REGION Network 6: Span Adjustment
   // Zero adjustment has to be performed prior to this linearity adjustment procedure.
   // 
   // 1. Specify how many linearity adjustment points to be performed by loading interger 0, 1, 2 or 3 into LinearityRange (0 for 2 points, 1 for 3 points, 2 for 4 points and 3 for 5 points). Please be noted that the earlier performed zero adjustment point is considered as the first adjustment point (Point #1).
   // 
   // 2. Configure all the adjustment weight values into xLow, Low, Middle and High (for e.g. 5-point adjustment requires all 4 weights: High, Middle, Low and xLow; 3-point requires High and Middle; 2-point only requies High as the 1st point is the zero reference)
   // 
   // 3. Make sure the Linearity Range parameter and all the adjustment weight values are configured correctly before starting the adjustment process. Invalid or incomplete parameters will cause the Function Block to turn on the Error output bit.
   // 
   // 4. Trigger ON  Input Start bit to start the span adjustment. This Start bit will be turned off by the Function Block upon completion/ cancellation or error condition. 
   // 
   // 5. Once started, CurrentPoint shows the current linearity point to be adjusted; CurrentWeight shows current adjustment weight to be loaded onto the scale. The LoadWeight output bit will be set ON to request for new adjustment weight. 
   // 
   // 6. After loading the new adjustment weight, acknowledge this by triggering the ConfirmWeight parameter (boolean) ON. The Function Block will then proceed to the next adjustment point and turn off this ConfirmWeight bit.
   // 
   // 7. Output bit - Process signifies that the adjustment of current point is in process.
   // 
   // 8. Input Parameter Bit Cancel is used to cancel/ abort the adjustment process
   RUNG wire#powerrail
      "SAI_IND_SpanAdjust_DB"(ID := "IND360~Head", Hi_Weight := "SAI_IND_SpanAdjust_DB".Hi_Weight, Mid_Weight := "SAI_IND_SpanAdjust_DB".Mid_Weight, Low_Weight := "SAI_IND_SpanAdjust_DB".Low_Weight, xLow_Weight := "SAI_IND_SpanAdjust_DB".xLow_Weight, LinearityRange := "SAI_IND_SpanAdjust_DB".LinearityRange, Start := "SAI_IND_SpanAdjust_DB".Start, ConfirmWeight := "SAI_IND_SpanAdjust_DB".ConfirmWeight, Cancel := "SAI_IND_SpanAdjust_DB".Cancel, CurrentPoint => "SAI_IND_SpanAdjust_DB".CurrentPoint, CurrentWeight => "SAI_IND_SpanAdjust_DB".CurrentWeight, LoadWeight => "SAI_IND_SpanAdjust_DB".LoadWeight, Process => "SAI_IND_SpanAdjust_DB".Process, Done => "SAI_IND_SpanAdjust_DB".Done, Error => "SAI_IND_SpanAdjust_DB".Error, Cancelled => "SAI_IND_SpanAdjust_DB".Cancelled)
   END_RUNG
   // the same network as SCL:
   "SAI_IND_SpanAdjust_DB"(ID := "IND360~Head",   // "SAI_IND_SpanAdjust"
                           Hi_Weight := "SAI_IND_SpanAdjust_DB".Hi_Weight,
                           Mid_Weight := "SAI_IND_SpanAdjust_DB".Mid_Weight,
                           Low_Weight := "SAI_IND_SpanAdjust_DB".Low_Weight,
                           xLow_Weight := "SAI_IND_SpanAdjust_DB".xLow_Weight,
                           LinearityRange := "SAI_IND_SpanAdjust_DB".LinearityRange,
                           Start := "SAI_IND_SpanAdjust_DB".Start,
                           ConfirmWeight := "SAI_IND_SpanAdjust_DB".ConfirmWeight,
                           Cancel := "SAI_IND_SpanAdjust_DB".Cancel,
                           CurrentPoint => "SAI_IND_SpanAdjust_DB".CurrentPoint,
                           CurrentWeight => "SAI_IND_SpanAdjust_DB".CurrentWeight,
                           LoadWeight => "SAI_IND_SpanAdjust_DB".LoadWeight,
                           Process => "SAI_IND_SpanAdjust_DB".Process,
                           Done => "SAI_IND_SpanAdjust_DB".Done,
                           Error => "SAI_IND_SpanAdjust_DB".Error,
                           Cancelled => "SAI_IND_SpanAdjust_DB".Cancelled);
END_REGION

REGION Network 7: CalFree Adjustment
   // CalFree is a method of analog scale adjustment without using test weights. It takes the factory calibrated load cell Rated Output (mV/ Vexc.) and user defined scale capacity to build a linear loading curve.
   // This method is usually applied to huge capacity scales in which calibration with test weights or other material is not feasible at all. 
   // 
   // For Powercell scale, please use the CalFree+ Function Block instead.
   // 
   // 1. Write in.. 
   // (a) CalFree Scale Capacity (Index 0x401A), 
   // (b) CalFree Scale unit (Index 0x401C, Decimal 0 - gram; Decimal 1 - KG; Decimal 2 - Pounds) and 
   // (c) Load Cells' averaged Rated Output (Index 0x401D, in mV/V)
   // **Make sure the transmitter's scale capacity has already been configured to the same value as CalFree Capacity prior to this CalFree adjustment.
   // 
   // 2. Trigger Input bit Start for CalFree adjustment (Index 0x401A)
   // 
   // 3. Output bit Done will be turned ON after successful completion of the process
   // Error output bit will be turned ON if there is an error during the adjustment process
   RUNG wire#powerrail
      "SAI_IND_CalFree_DB"(ID := "IND360~Head", RatedCapacity := "SAI_IND_CalFree_DB".RatedCapacity, Unit := "SAI_IND_CalFree_DB".Unit, RatedOutput := "SAI_IND_CalFree_DB".RatedOutput, Start := "SAI_IND_CalFree_DB".Start, Process => "SAI_IND_CalFree_DB".Process, Done => "SAI_IND_CalFree_DB".Done, Error => "SAI_IND_CalFree_DB".Error)
   END_RUNG
   // the same network as SCL:
   "SAI_IND_CalFree_DB"(ID := "IND360~Head",   // "SAI_IND_CalFree"
                        RatedCapacity := "SAI_IND_CalFree_DB".RatedCapacity,
                        Unit := "SAI_IND_CalFree_DB".Unit,
                        RatedOutput := "SAI_IND_CalFree_DB".RatedOutput,
                        Start := "SAI_IND_CalFree_DB".Start,
                        Process => "SAI_IND_CalFree_DB".Process,
                        Done => "SAI_IND_CalFree_DB".Done,
                        Error => "SAI_IND_CalFree_DB".Error);
END_REGION

REGION Network 8: Alibi Record Read
   // Use this Function Block to read one alibi record. 
   // 1. Set the alibi transaction number to be read.
   // 2. Toggle the Get_Record bit to perform read. Alibi record will be written into Alibi_Array (an array of 44 Bytes).  
   // 3. The read alibi record transaction gross, net and tare weights (all LREAL format) as well as weight unit are available at the FB's output.
   // 4. the Alibi_Array structure data format is as below:
   // 
   // For Base, RateControl, Tank Vessel:
   // Struct(44 Bytes)
   // {
   // Byte[20]: Date & time; //ASCII String  =>Byte0-19
   // Long:     Transaction Number;            =>Byte20-23
   // Float32:  Gross Weight;                       =>Byte24-27
   // Float32:  Net Weight;                           =>Byte28-31
   // Float32:  Tare Weight;                         =>Byte32-35
   // Byte:     Tare Mode;                              =>Byte36
   // Byte:     Unit;                                          =>Byte37
   // Byte[6]:  Not Used;                              =>Byte38-43
   // }
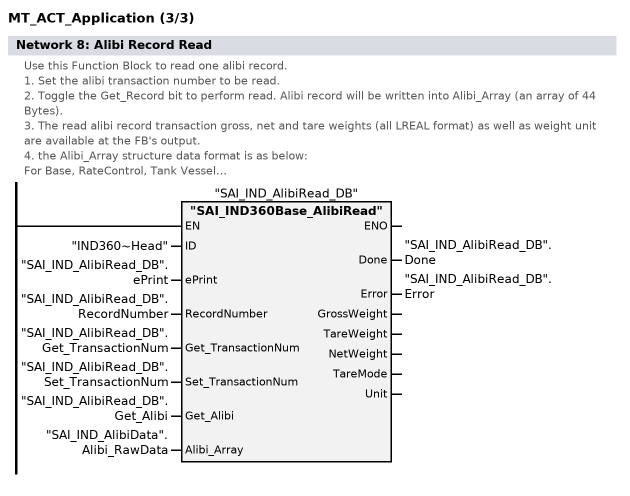
   RUNG wire#powerrail
      "SAI_IND_AlibiRead_DB"(ID := "IND360~Head", ePrint := "SAI_IND_AlibiRead_DB".ePrint, RecordNumber := "SAI_IND_AlibiRead_DB".RecordNumber, Get_TransactionNum := "SAI_IND_AlibiRead_DB".Get_TransactionNum, Set_TransactionNum := "SAI_IND_AlibiRead_DB".Set_TransactionNum, Get_Alibi := "SAI_IND_AlibiRead_DB".Get_Alibi, Alibi_Array := "SAI_IND_AlibiData".Alibi_RawData, Done => "SAI_IND_AlibiRead_DB".Done, Error => "SAI_IND_AlibiRead_DB".Error, GrossWeight =>, TareWeight =>, NetWeight =>, TareMode =>, Unit =>)
   END_RUNG
   // the same network as SCL:
   "SAI_IND_AlibiRead_DB"(ID := "IND360~Head",   // "SAI_IND360Base_AlibiRead"
                          ePrint := "SAI_IND_AlibiRead_DB".ePrint,
                          RecordNumber := "SAI_IND_AlibiRead_DB".RecordNumber,
                          Get_TransactionNum := "SAI_IND_AlibiRead_DB".Get_TransactionNum,
                          Set_TransactionNum := "SAI_IND_AlibiRead_DB".Set_TransactionNum,
                          Get_Alibi := "SAI_IND_AlibiRead_DB".Get_Alibi,
                          Alibi_Array := "SAI_IND_AlibiData".Alibi_RawData,
                          Done => "SAI_IND_AlibiRead_DB".Done,
                          Error => "SAI_IND_AlibiRead_DB".Error);
END_REGION
END_FUNCTION

FUNCTION_BLOCK "SAI_Cyclic_WeightProc"   // FB29, LAD
TITLE = Cyclic Weighing Process: Send PLC commands and read Weight data and device status bits
{ S7_Optimized_Access := 'FALSE' }
VERSION : 0.1
// stored: AutoNumber true, IsIECCheckEnabled false, SetENOAutomatically false, UDAEnableTagReadback false
   VAR_INPUT
      WeightCmd { ExternalAccessible := 'False'; ExternalVisible := 'False'; ExternalWritable := 'False'} : Word := 3;
      MB_DevStatus : Word;
   END_VAR
   VAR_OUTPUT
      RealTimeWeight { ExternalVisible := 'False'; ExternalWritable := 'False'} : Real;
      StableWeight { ExternalVisible := 'False'; ExternalWritable := 'False'} : Real;
      DataOK : Bool;
      Motion : Bool;
      NetMode : Bool;
      Alarm : Bool;
      Done { ExternalAccessible := 'False'; ExternalVisible := 'False'; ExternalWritable := 'False'} : Bool;
      Error { ExternalAccessible := 'False'; ExternalVisible := 'False'; ExternalWritable := 'False'} : Bool;
   END_VAR
   VAR_IN_OUT
      TareImmediate { ExternalAccessible := 'False'; ExternalVisible := 'False'; ExternalWritable := 'False'} : Bool;
      TareStable { ExternalAccessible := 'False'; ExternalVisible := 'False'; ExternalWritable := 'False'} : Bool;
      ZeroImmediate { ExternalAccessible := 'False'; ExternalVisible := 'False'; ExternalWritable := 'False'} : Bool;
      ZeroStable { ExternalAccessible := 'False'; ExternalVisible := 'False'; ExternalWritable := 'False'} : Bool;
      PreTareValue : Real;
      PreTare : Bool;
      ClearTare { ExternalAccessible := 'False'; ExternalVisible := 'False'; ExternalWritable := 'False'} : Bool;
      MB_Value : Real;
      MB_Response : Word;
      MB_CmdValue : Real;
      MB_Command : Word;
   END_VAR
   VAR DB_SPECIFIC
      WriteTrigger { ExternalAccessible := 'False'; ExternalVisible := 'False'; ExternalWritable := 'False'} : Bool;
      RestoreTrigger { ExternalAccessible := 'False'; ExternalVisible := 'False'; ExternalWritable := 'False'} : Bool;
      Cmd { ExternalAccessible := 'False'; ExternalVisible := 'False'; ExternalWritable := 'False'} : Int;
      TareStablePTrigger : Bool;
      ZeroStablePTrigger : Bool;
      ZeroImmedTrigger : Bool;
      TareImmedTrigger : Bool;
      ClearTareTrigger : Bool;
      PreTareTrigger : Bool;
   END_VAR
   VAR_TEMP
      DevStatus : "SAI_MB_DeviceStatus";
   END_VAR
   VAR_TEMP   // added for the SCL form of the ladder/FBD networks
      _w1 : Bool;
   END_VAR
BEGIN

REGION Network 1: During 1st PLC scan, moves the default weight reporting command to the cyclic command output word
   // During 1st scan, moves the default weight reporting command to the cyclic command output word
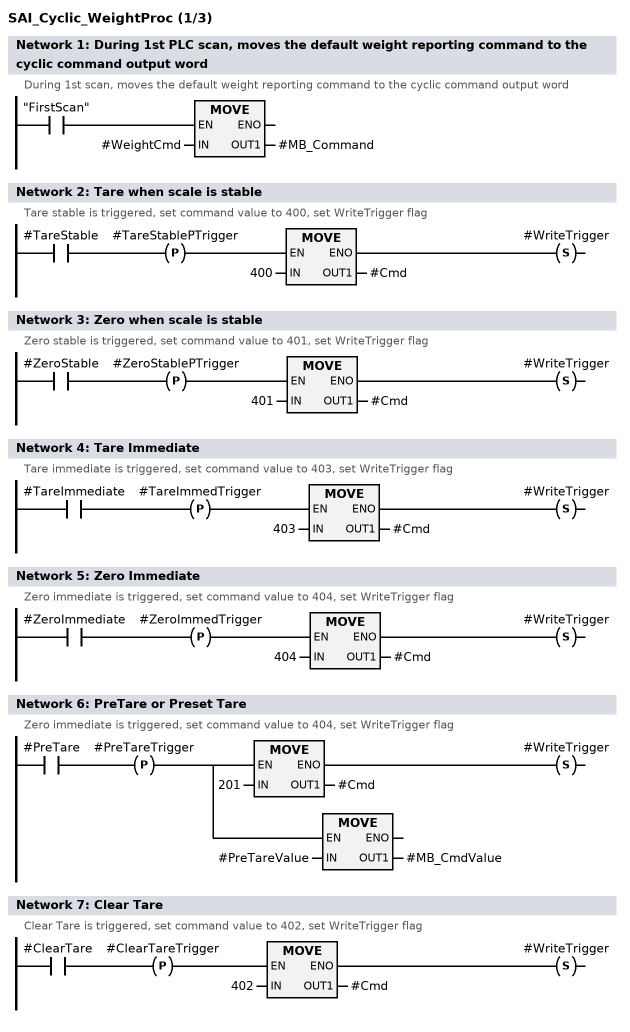
   RUNG wire#powerrail
      Contact( "FirstScan" )
      { S7_GenerateENO := "TRUE" } Move(in := #WeightCmd, out1 => #MB_Command)
   END_RUNG
   // the same network as SCL:
   IF "FirstScan" THEN #MB_Command := #WeightCmd; END_IF;
END_REGION

REGION Network 2: Tare when scale is stable
   // Tare stable is triggered, set command value to 400, set WriteTrigger flag
   RUNG wire#powerrail
      Contact( #TareStable )
      P_Trig( #TareStablePTrigger )
      { S7_GenerateENO := "TRUE" } Move(in := 400, out1 => #Cmd)
      S_Coil( #WriteTrigger )
   END_RUNG
   // the same network as SCL:
   // ENO of a box is taken as its EN; it also drops when the box reports an error
   #_w1 := #TareStable AND NOT #TareStablePTrigger;   // rising edge
   #TareStablePTrigger := #TareStable;
   IF #_w1 THEN
       #Cmd := 400;
       #WriteTrigger := TRUE;
   END_IF;
END_REGION

REGION Network 3: Zero when scale is stable
   // Zero stable is triggered, set command value to 401, set WriteTrigger flag
   RUNG wire#powerrail
      Contact( #ZeroStable )
      P_Trig( #ZeroStablePTrigger )
      { S7_GenerateENO := "TRUE" } Move(in := 401, out1 => #Cmd)
      S_Coil( #WriteTrigger )
   END_RUNG
   // the same network as SCL:
   // ENO of a box is taken as its EN; it also drops when the box reports an error
   #_w1 := #ZeroStable AND NOT #ZeroStablePTrigger;   // rising edge
   #ZeroStablePTrigger := #ZeroStable;
   IF #_w1 THEN
       #Cmd := 401;
       #WriteTrigger := TRUE;
   END_IF;
END_REGION

REGION Network 4: Tare Immediate
   // Tare immediate is triggered, set command value to 403, set WriteTrigger flag
   RUNG wire#powerrail
      Contact( #TareImmediate )
      P_Trig( #TareImmedTrigger )
      { S7_GenerateENO := "TRUE" } Move(in := 403, out1 => #Cmd)
      S_Coil( #WriteTrigger )
   END_RUNG
   // the same network as SCL:
   // ENO of a box is taken as its EN; it also drops when the box reports an error
   #_w1 := #TareImmediate AND NOT #TareImmedTrigger;   // rising edge
   #TareImmedTrigger := #TareImmediate;
   IF #_w1 THEN
       #Cmd := 403;
       #WriteTrigger := TRUE;
   END_IF;
END_REGION

REGION Network 5: Zero Immediate
   // Zero immediate is triggered, set command value to 404, set WriteTrigger flag
   RUNG wire#powerrail
      Contact( #ZeroImmediate )
      P_Trig( #ZeroImmedTrigger )
      { S7_GenerateENO := "TRUE" } Move(in := 404, out1 => #Cmd)
      S_Coil( #WriteTrigger )
   END_RUNG
   // the same network as SCL:
   // ENO of a box is taken as its EN; it also drops when the box reports an error
   #_w1 := #ZeroImmediate AND NOT #ZeroImmedTrigger;   // rising edge
   #ZeroImmedTrigger := #ZeroImmediate;
   IF #_w1 THEN
       #Cmd := 404;
       #WriteTrigger := TRUE;
   END_IF;
END_REGION

REGION Network 6: PreTare or Preset Tare
   // Zero immediate is triggered, set command value to 404, set WriteTrigger flag
   RUNG wire#powerrail
      Contact( #PreTare )
      P_Trig( #PreTareTrigger )
      wire#w1
      { S7_GenerateENO := "TRUE" } Move(in := 201, out1 => #Cmd)
      S_Coil( #WriteTrigger )
   END_RUNG
   RUNG wire#w1
      { S7_GenerateENO := "TRUE" } Move(in := #PreTareValue, out1 => #MB_CmdValue)
   END_RUNG
   // the same network as SCL:
   // ENO of a box is taken as its EN; it also drops when the box reports an error
   #_w1 := #PreTare AND NOT #PreTareTrigger;   // rising edge
   #PreTareTrigger := #PreTare;
   IF #_w1 THEN
       #Cmd := 201;
       #WriteTrigger := TRUE;
       #MB_CmdValue := #PreTareValue;
   END_IF;
END_REGION

REGION Network 7: Clear Tare
   // Clear Tare is triggered, set command value to 402, set WriteTrigger flag
   RUNG wire#powerrail
      Contact( #ClearTare )
      P_Trig( #ClearTareTrigger )
      { S7_GenerateENO := "TRUE" } Move(in := 402, out1 => #Cmd)
      S_Coil( #WriteTrigger )
   END_RUNG
   // the same network as SCL:
   // ENO of a box is taken as its EN; it also drops when the box reports an error
   #_w1 := #ClearTare AND NOT #ClearTareTrigger;   // rising edge
   #ClearTareTrigger := #ClearTare;
   IF #_w1 THEN
       #Cmd := 402;
       #WriteTrigger := TRUE;
   END_IF;
END_REGION

REGION Network 8: Deliver the command
   // Move the command value to output, reset flags
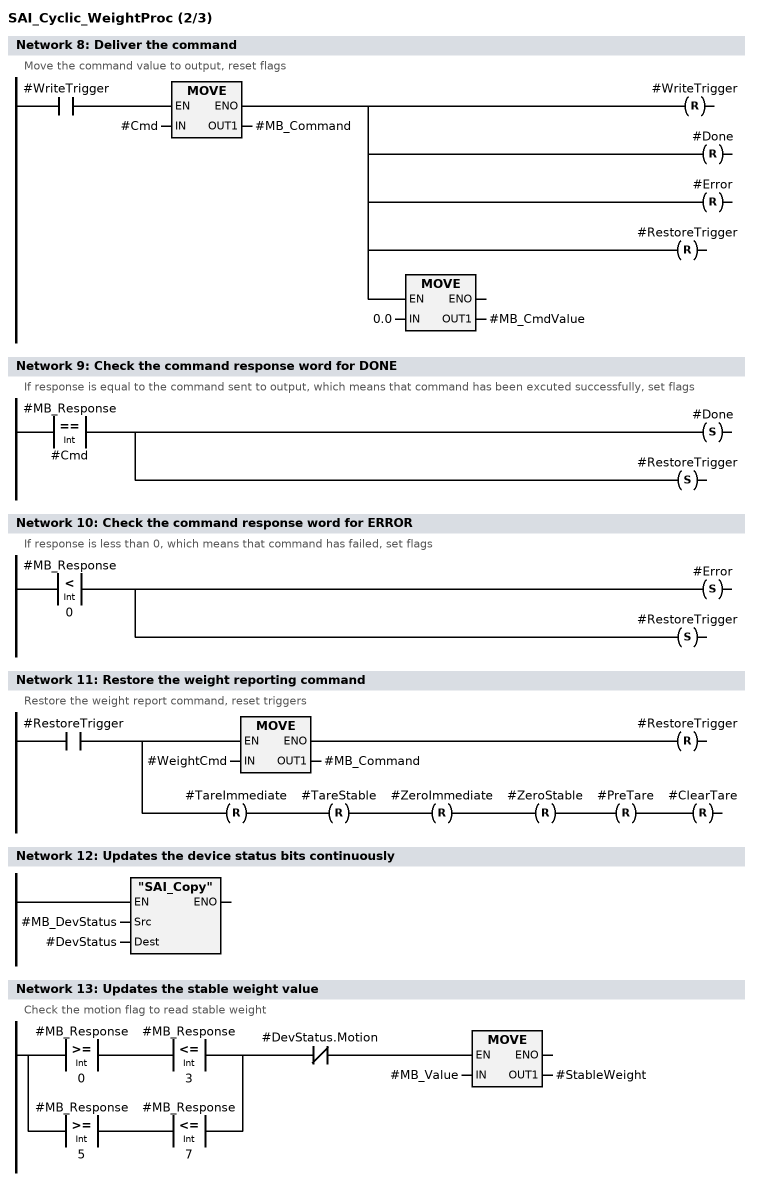
   RUNG wire#powerrail
      Contact( #WriteTrigger )
      { S7_GenerateENO := "TRUE" } Move(in := #Cmd, out1 => #MB_Command)
      wire#w1
      R_Coil( #WriteTrigger )
   END_RUNG
   RUNG wire#w1
      R_Coil( #Done )
   END_RUNG
   RUNG wire#w1
      R_Coil( #Error )
   END_RUNG
   RUNG wire#w1
      R_Coil( #RestoreTrigger )
   END_RUNG
   RUNG wire#w1
      { S7_GenerateENO := "TRUE" } Move(in := 0.0, out1 => #MB_CmdValue)
   END_RUNG
   // the same network as SCL:
   // ENO of a box is taken as its EN; it also drops when the box reports an error
   IF #WriteTrigger THEN #MB_Command := #Cmd; END_IF;
   #_w1 := #WriteTrigger;
   IF #_w1 THEN
       #WriteTrigger := FALSE;
       #Done := FALSE;
       #Error := FALSE;
       #RestoreTrigger := FALSE;
       #MB_CmdValue := 0.0;
   END_IF;
END_REGION

REGION Network 9: Check the command response word for DONE
   // If response is equal to the command sent to output, which means that command has been excuted successfully, set flags
   RUNG wire#powerrail
      { S7_Templates := "SrcType := Int" } EQ_Contact(in1 := #MB_Response, in2 := #Cmd)
      wire#w1
      S_Coil( #Done )
   END_RUNG
   RUNG wire#w1
      S_Coil( #RestoreTrigger )
   END_RUNG
   // the same network as SCL:
   IF #MB_Response = #Cmd THEN
       #Done := TRUE;
       #RestoreTrigger := TRUE;
   END_IF;
END_REGION

REGION Network 10: Check the command response word for ERROR
   // If response is less than 0, which means that command has failed, set flags
   RUNG wire#powerrail
      { S7_Templates := "SrcType := Int" } LT_Contact(in1 := #MB_Response, in2 := 0)
      wire#w1
      S_Coil( #Error )
   END_RUNG
   RUNG wire#w1
      S_Coil( #RestoreTrigger )
   END_RUNG
   // the same network as SCL:
   IF #MB_Response < 0 THEN
       #Error := TRUE;
       #RestoreTrigger := TRUE;
   END_IF;
END_REGION

REGION Network 11: Restore the weight reporting command
   // Restore the weight report command, reset triggers
   RUNG wire#powerrail
      Contact( #RestoreTrigger )
      wire#w1
      { S7_GenerateENO := "TRUE" } Move(in := #WeightCmd, out1 => #MB_Command)
      R_Coil( #RestoreTrigger )
   END_RUNG
   RUNG wire#w1
      R_Coil( #TareImmediate )
      R_Coil( #TareStable )
      R_Coil( #ZeroImmediate )
      R_Coil( #ZeroStable )
      R_Coil( #PreTare )
      R_Coil( #ClearTare )
   END_RUNG
   // the same network as SCL:
   // ENO of a box is taken as its EN; it also drops when the box reports an error
   IF #RestoreTrigger THEN #MB_Command := #WeightCmd; END_IF;
   #_w1 := #RestoreTrigger;
   IF #_w1 THEN
       #RestoreTrigger := FALSE;
       #TareImmediate := FALSE;
       #TareStable := FALSE;
       #ZeroImmediate := FALSE;
       #ZeroStable := FALSE;
       #PreTare := FALSE;
       #ClearTare := FALSE;
   END_IF;
END_REGION

REGION Network 12: Updates the device status bits continuously
   RUNG wire#powerrail
      "SAI_Copy"(Src := #MB_DevStatus, Dest := #DevStatus)
   END_RUNG
   // the same network as SCL:
   "SAI_Copy"(Src := #MB_DevStatus, Dest := #DevStatus);
END_REGION

REGION Network 13: Updates the stable weight value
   // Check the motion flag to read stable weight
   RUNG wire#powerrail
      { S7_Templates := "SrcType := Int" } GE_Contact(in1 := #MB_Response, in2 := 0)
      { S7_Templates := "SrcType := Int" } LE_Contact(in1 := #MB_Response, in2 := 3)
      wire#w1
      I_Contact( #DevStatus.Motion )
      { S7_GenerateENO := "TRUE" } Move(in := #MB_Value, out1 => #StableWeight)
   END_RUNG
   RUNG wire#powerrail
      { S7_Templates := "SrcType := Int" } GE_Contact(in1 := #MB_Response, in2 := 5)
      { S7_Templates := "SrcType := Int" } LE_Contact(in1 := #MB_Response, in2 := 7)
   END_RUNG wire#w1
   // the same network as SCL:
   IF (((#MB_Response >= 0) AND (#MB_Response <= 3)) OR ((#MB_Response >= 5) AND (#MB_Response <= 7))) AND NOT #DevStatus.Motion THEN
       #StableWeight := #MB_Value;
   END_IF;
END_REGION

REGION Network 14: Updates the real time weight value
   // Read real time weight
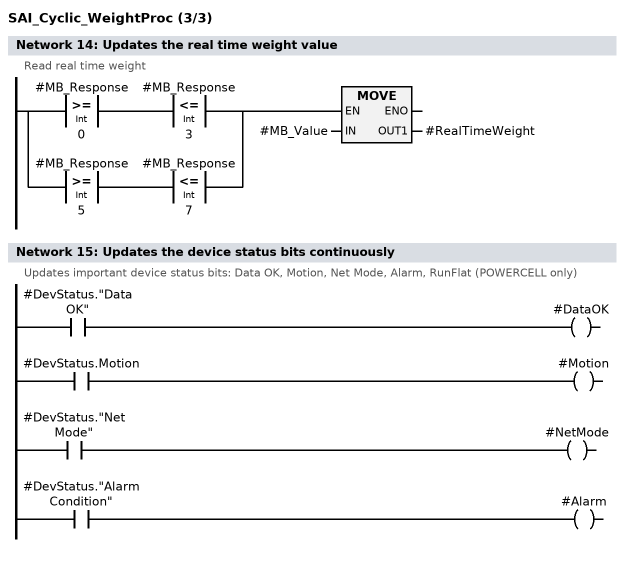
   RUNG wire#powerrail
      { S7_Templates := "SrcType := Int" } GE_Contact(in1 := #MB_Response, in2 := 0)
      { S7_Templates := "SrcType := Int" } LE_Contact(in1 := #MB_Response, in2 := 3)
      wire#w1
      { S7_GenerateENO := "TRUE" } Move(in := #MB_Value, out1 => #RealTimeWeight)
   END_RUNG
   RUNG wire#powerrail
      { S7_Templates := "SrcType := Int" } GE_Contact(in1 := #MB_Response, in2 := 5)
      { S7_Templates := "SrcType := Int" } LE_Contact(in1 := #MB_Response, in2 := 7)
   END_RUNG wire#w1
   // the same network as SCL:
   IF ((#MB_Response >= 0) AND (#MB_Response <= 3)) OR ((#MB_Response >= 5) AND (#MB_Response <= 7)) THEN
       #RealTimeWeight := #MB_Value;
   END_IF;
END_REGION

REGION Network 15: Updates the device status bits continuously
   // Updates important device status bits: Data OK, Motion, Net Mode, Alarm, RunFlat (POWERCELL only)
   RUNG wire#powerrail
      Contact( #DevStatus."Data OK" )
      Coil( #DataOK )
   END_RUNG
   RUNG wire#powerrail
      Contact( #DevStatus.Motion )
      Coil( #Motion )
   END_RUNG
   RUNG wire#powerrail
      Contact( #DevStatus."Net Mode" )
      Coil( #NetMode )
   END_RUNG
   RUNG wire#powerrail
      Contact( #DevStatus."Alarm Condition" )
      Coil( #Alarm )
   END_RUNG
   // the same network as SCL:
   #DataOK := #DevStatus."Data OK";
   #Motion := #DevStatus.Motion;
   #NetMode := #DevStatus."Net Mode";
   #Alarm := #DevStatus."Alarm Condition";
END_REGION
END_FUNCTION_BLOCK

FUNCTION "SAI_Copy" : Void   // FC29, LAD
{ S7_Optimized_Access := 'FALSE' }
VERSION : 0.1
// stored: AutoNumber true, IsIECCheckEnabled false, SetENOAutomatically false, UDAEnableTagReadback false
   VAR_INPUT
      Src : Variant;
   END_VAR
   VAR_IN_OUT
      Dest : Variant;
   END_VAR
   VAR_TEMP
      TmpBuf : Array[0..100] of Byte;
      TmpRet : Int;
      TmpPos : DInt;
   END_VAR
BEGIN

REGION Network 1
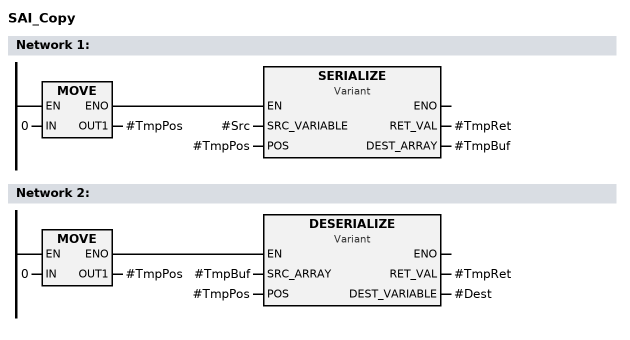
   RUNG wire#powerrail
      Move(in := 0, out1 => #TmpPos)
      { S7_Templates := "[src_type := Variant, dest_type := Variant]" } Serialize(SRC_VARIABLE := #Src, POS := #TmpPos, Ret_Val => #TmpRet, DEST_ARRAY => #TmpBuf)
   END_RUNG
   // the same network as SCL:
   #TmpPos := 0;
   #TmpRet := Serialize(SRC_VARIABLE := #Src, POS := #TmpPos, DEST_ARRAY => #TmpBuf);
END_REGION

REGION Network 2
   RUNG wire#powerrail
      Move(in := 0, out1 => #TmpPos)
      { S7_Templates := "[src_type := Variant, dest_type := Variant]" } Deserialize(SRC_ARRAY := #TmpBuf, POS := #TmpPos, Ret_Val => #TmpRet, DEST_VARIABLE => #Dest)
   END_RUNG
   // the same network as SCL:
   #TmpPos := 0;
   #TmpRet := Deserialize(SRC_ARRAY := #TmpBuf, POS := #TmpPos, DEST_VARIABLE => #Dest);
END_REGION
END_FUNCTION

FUNCTION_BLOCK "SAI_Cyclic_CheckAlive"   // FB28, LAD
TITLE = Check HearBeat status bit and update the Alive bit
{ S7_Optimized_Access := 'FALSE' }
VERSION : 0.1
// stored: AutoNumber true, IsIECCheckEnabled false, SetENOAutomatically false, UDAEnableTagReadback false
   VAR_INPUT
      MB_DevStatus : Word;
   END_VAR
   VAR_OUTPUT
      Alive : Bool;
      HeartBeat : Bool;
   END_VAR
   VAR DB_SPECIFIC
      PTrigHeart : Bool;
      NTrigHeart : Bool;
      bResetTimer : Bool;
      IEC_Timer { S7_SetPoint := 'True'} : IEC_TIMER;
   END_VAR
   VAR_TEMP
      DevStatus : "SAI_MB_DeviceStatus";
   END_VAR
   VAR_TEMP   // added for the SCL form of the ladder/FBD networks
      _w1 : Bool;
      _w2 : Bool;
      _w3 : Bool;
   END_VAR
BEGIN

REGION Network 1: Gets the cyclic device status - HeartBeat bit
   // Gets the cyclic device status - HeartBeat bit
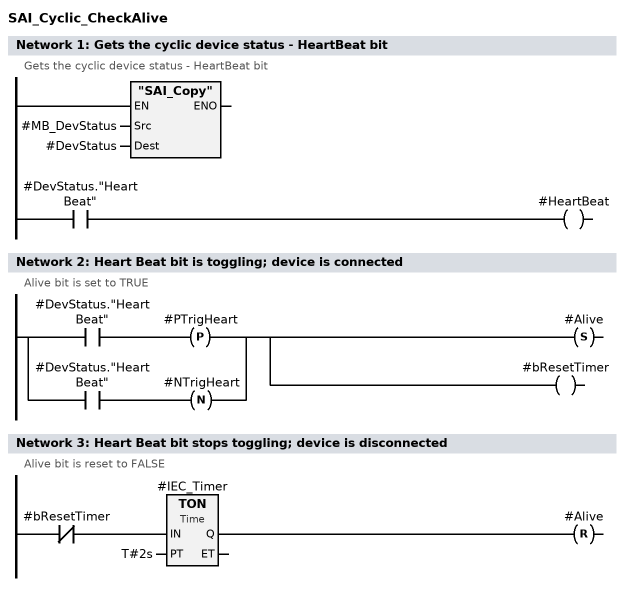
   RUNG wire#powerrail
      "SAI_Copy"(Src := #MB_DevStatus, Dest := #DevStatus)
   END_RUNG
   RUNG wire#powerrail
      Contact( #DevStatus."Heart Beat" )
      Coil( #HeartBeat )
   END_RUNG
   // the same network as SCL:
   "SAI_Copy"(Src := #MB_DevStatus, Dest := #DevStatus);
   #HeartBeat := #DevStatus."Heart Beat";
END_REGION

REGION Network 2: Heart Beat bit is toggling; device is connected
   // Alive bit is set to TRUE
   RUNG wire#powerrail
      Contact( #DevStatus."Heart Beat" )
      P_Trig( #PTrigHeart )
      wire#w1
      S_Coil( #Alive )
   END_RUNG
   RUNG wire#powerrail
      Contact( #DevStatus."Heart Beat" )
      N_Trig( #NTrigHeart )
   END_RUNG wire#w1
   RUNG wire#w1
      Coil( #bResetTimer )
   END_RUNG
   // the same network as SCL:
   #_w1 := #DevStatus."Heart Beat" AND NOT #PTrigHeart;   // rising edge
   #PTrigHeart := #DevStatus."Heart Beat";
   #_w2 := NOT #DevStatus."Heart Beat" AND #NTrigHeart;   // falling edge
   #NTrigHeart := #DevStatus."Heart Beat";
   #_w3 := #_w1 OR #_w2;
   IF #_w3 THEN #Alive := TRUE; END_IF;
   #bResetTimer := #_w3;
END_REGION

REGION Network 3: Heart Beat bit stops toggling; device is disconnected
   // Alive bit is reset to FALSE
   RUNG wire#powerrail
      I_Contact( #bResetTimer )
      { S7_Templates := "time_type := Time" } #IEC_Timer.TON(pt := T#2s, et =>)
      R_Coil( #Alive )
   END_RUNG
   // the same network as SCL:
   #IEC_Timer.TON(IN := NOT #bResetTimer, PT := T#2s);
   IF #IEC_Timer.Q THEN #Alive := FALSE; END_IF;
END_REGION
END_FUNCTION_BLOCK

FUNCTION_BLOCK "SAI_IND_ReadAdjustSettings"   // FB50, LAD
{ S7_Optimized_Access := 'FALSE' }
VERSION : 0.1
// stored: AutoNumber true, IsIECCheckEnabled false, SetENOAutomatically false, UDAEnableTagReadback false
   VAR_INPUT
      ID : HW_IO;   // The Profinet Device Hardware Identifier under device properties
   END_VAR
   VAR_OUTPUT
      ScaleCapacity : Real;   // The configured scale capacity
      Increment : Real;   // The configured scale increment value
      Done : Bool;   // Read done successfully
      Error : Bool;   // Error during reading process
   END_VAR
   VAR_IN_OUT
      Read : Bool;   // Switch this bit ON to start reading
   END_VAR
   VAR DB_SPECIFIC
      Static01 : Bool;
      "Step" : Int;
   END_VAR
   VAR
      RDREC_CAP { S7_SetPoint := 'True'} : RDREC;
   END_VAR
   VAR DB_SPECIFIC
      CAP_RECORD : Real;
      INC_RECORD : Real;
      Activate : Bool;
   END_VAR
   VAR_TEMP
      Temp02 : Bool;
   END_VAR
   VAR_TEMP   // added for the SCL form of the ladder/FBD networks
      _w1 : Bool;
      _w2 : Bool;
      _w3 : Bool;
      _w4 : Bool;
      _w5 : Bool;
      _w6 : Bool;
      _w7 : Bool;
   END_VAR
BEGIN

REGION Network 1: Initialization
   // Initializes FB output bits:
   // Error;
   // Done;
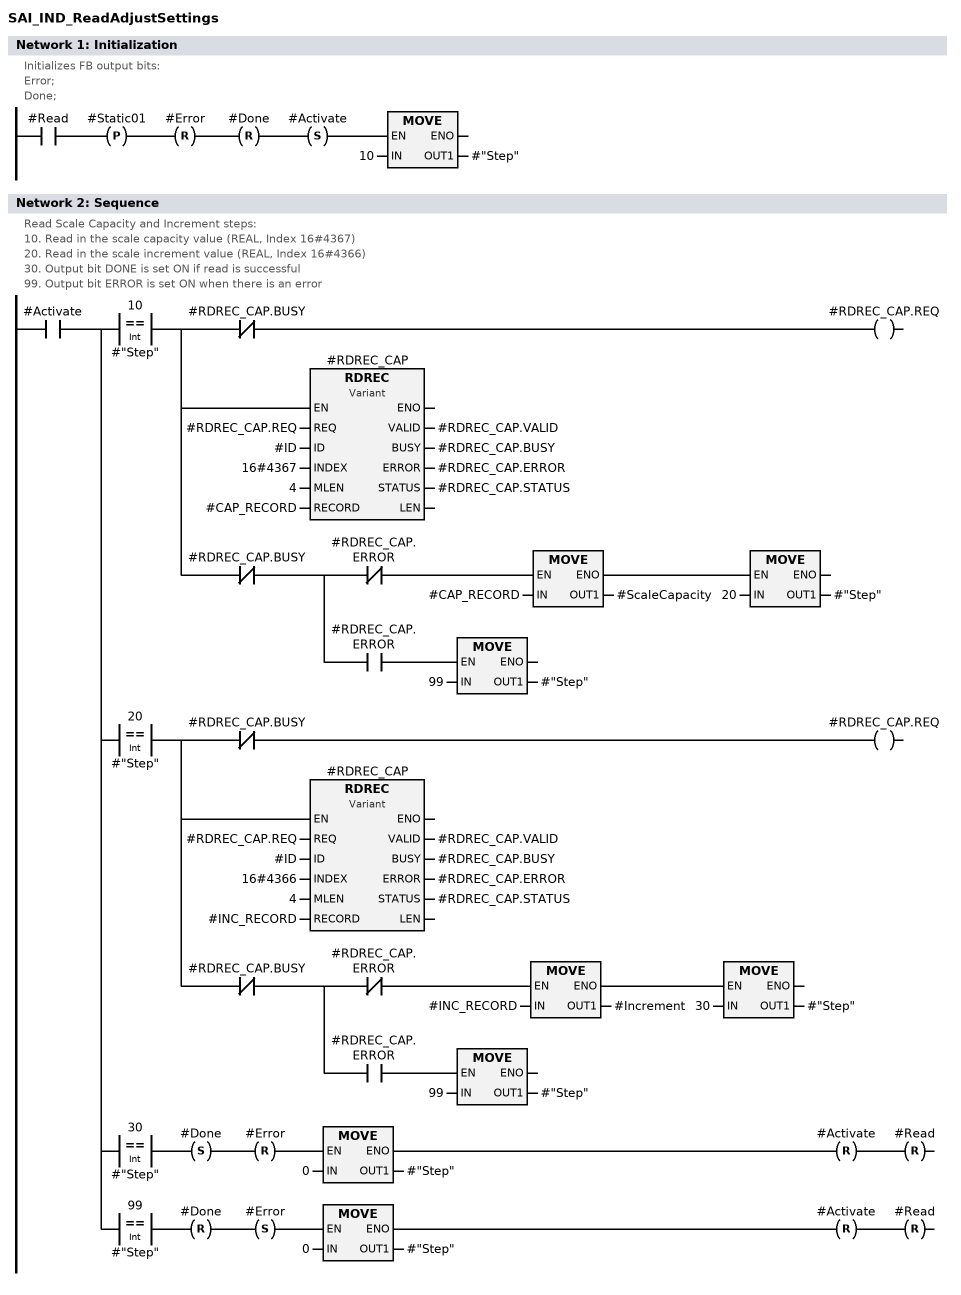
   RUNG wire#powerrail
      Contact( #Read )
      P_Trig( #Static01 )
      R_Coil( #Error )
      R_Coil( #Done )
      S_Coil( #Activate )
      { S7_GenerateENO := "TRUE" } Move(in := 10, out1 => #"Step")
   END_RUNG
   // the same network as SCL:
   #_w1 := #Read AND NOT #Static01;   // rising edge
   #Static01 := #Read;
   IF #_w1 THEN
       #Error := FALSE;
       #Done := FALSE;
       #Activate := TRUE;
       #"Step" := 10;
   END_IF;
END_REGION

REGION Network 2: Sequence
   // Read Scale Capacity and Increment steps:
   // 10. Read in the scale capacity value (REAL, Index 16#4367) 
   // 20. Read in the scale increment value (REAL, Index 16#4366) 
   // 30. Output bit DONE is set ON if read is successful
   // 99. Output bit ERROR is set ON when there is an error
   RUNG wire#powerrail
      Contact( #Activate )
      wire#w1
      { S7_Templates := "SrcType := Int" } EQ_Contact(in1 := 10, in2 := #"Step")
      wire#w2
      I_Contact( #RDREC_CAP.BUSY )
      Coil( #RDREC_CAP.REQ )
   END_RUNG
   RUNG wire#w2
      { S7_Templates := "[ptr_type := Variant, id_type := HW_IO, index_type := DInt, len_type := UInt]" } #RDREC_CAP.RDREC(REQ := #RDREC_CAP.REQ, ID := #ID, INDEX := 16#4367, MLEN := 4, RECORD := #CAP_RECORD, VALID => #RDREC_CAP.VALID, BUSY => #RDREC_CAP.BUSY, ERROR => #RDREC_CAP.ERROR, STATUS => #RDREC_CAP.STATUS, LEN =>)
   END_RUNG
   RUNG wire#w2
      I_Contact( #RDREC_CAP.BUSY )
      wire#w3
      I_Contact( #RDREC_CAP.ERROR )
      { S7_GenerateENO := "TRUE" } Move(in := #CAP_RECORD, out1 => #ScaleCapacity)
      { S7_GenerateENO := "TRUE" } Move(in := 20, out1 => #"Step")
   END_RUNG
   RUNG wire#w3
      Contact( #RDREC_CAP.ERROR )
      { S7_GenerateENO := "TRUE" } Move(in := 99, out1 => #"Step")
   END_RUNG
   RUNG wire#w1
      { S7_Templates := "SrcType := Int" } EQ_Contact(in1 := 20, in2 := #"Step")
      wire#w4
      I_Contact( #RDREC_CAP.BUSY )
      Coil( #RDREC_CAP.REQ )
   END_RUNG
   RUNG wire#w4
      { S7_Templates := "[ptr_type := Variant, id_type := HW_IO, index_type := DInt, len_type := UInt]" } #RDREC_CAP.RDREC(REQ := #RDREC_CAP.REQ, ID := #ID, INDEX := 16#4366, MLEN := 4, RECORD := #INC_RECORD, VALID => #RDREC_CAP.VALID, BUSY => #RDREC_CAP.BUSY, ERROR => #RDREC_CAP.ERROR, STATUS => #RDREC_CAP.STATUS, LEN =>)
   END_RUNG
   RUNG wire#w4
      I_Contact( #RDREC_CAP.BUSY )
      wire#w5
      I_Contact( #RDREC_CAP.ERROR )
      { S7_GenerateENO := "TRUE" } Move(in := #INC_RECORD, out1 => #Increment)
      { S7_GenerateENO := "TRUE" } Move(in := 30, out1 => #"Step")
   END_RUNG
   RUNG wire#w5
      Contact( #RDREC_CAP.ERROR )
      { S7_GenerateENO := "TRUE" } Move(in := 99, out1 => #"Step")
   END_RUNG
   RUNG wire#w1
      { S7_Templates := "SrcType := Int" } EQ_Contact(in1 := 30, in2 := #"Step")
      S_Coil( #Done )
      R_Coil( #Error )
      { S7_GenerateENO := "TRUE" } Move(in := 0, out1 => #"Step")
      R_Coil( #Activate )
      R_Coil( #Read )
   END_RUNG
   RUNG wire#w1
      { S7_Templates := "SrcType := Int" } EQ_Contact(in1 := 99, in2 := #"Step")
      R_Coil( #Done )
      S_Coil( #Error )
      { S7_GenerateENO := "TRUE" } Move(in := 0, out1 => #"Step")
      R_Coil( #Activate )
      R_Coil( #Read )
   END_RUNG
   // the same network as SCL:
   // ENO of a box is taken as its EN; it also drops when the box reports an error
   #_w1 := #Activate AND (10 = #"Step");
   #RDREC_CAP.REQ := #_w1 AND NOT #RDREC_CAP.BUSY;
   IF #_w1 THEN
       #RDREC_CAP(REQ := #RDREC_CAP.REQ,   // RDREC
                  ID := #ID,
                  INDEX := 16#4367,
                  MLEN := 4,
                  RECORD := #CAP_RECORD,
                  VALID => #RDREC_CAP.VALID,
                  BUSY => #RDREC_CAP.BUSY,
                  ERROR => #RDREC_CAP.ERROR,
                  STATUS => #RDREC_CAP.STATUS);
   END_IF;
   #_w2 := #_w1 AND NOT #RDREC_CAP.BUSY;
   IF #_w2 AND NOT #RDREC_CAP.ERROR THEN
       #ScaleCapacity := #CAP_RECORD;
       #"Step" := 20;
   END_IF;
   IF #_w2 AND #RDREC_CAP.ERROR THEN #"Step" := 99; END_IF;
   #_w3 := #Activate AND (20 = #"Step");
   #RDREC_CAP.REQ := #_w3 AND NOT #RDREC_CAP.BUSY;
   IF #_w3 THEN
       #RDREC_CAP(REQ := #RDREC_CAP.REQ,   // RDREC
                  ID := #ID,
                  INDEX := 16#4366,
                  MLEN := 4,
                  RECORD := #INC_RECORD,
                  VALID => #RDREC_CAP.VALID,
                  BUSY => #RDREC_CAP.BUSY,
                  ERROR => #RDREC_CAP.ERROR,
                  STATUS => #RDREC_CAP.STATUS);
   END_IF;
   #_w4 := #_w3 AND NOT #RDREC_CAP.BUSY;
   IF #_w4 AND NOT #RDREC_CAP.ERROR THEN
       #Increment := #INC_RECORD;
       #"Step" := 30;
   END_IF;
   IF #_w4 AND #RDREC_CAP.ERROR THEN #"Step" := 99; END_IF;
   IF #Activate AND (30 = #"Step") THEN
       #Done := TRUE;
       #Error := FALSE;
   END_IF;
   #_w5 := #Activate AND (30 = #"Step");
   IF #_w5 THEN #"Step" := 0; END_IF;
   #_w6 := #Activate;
   IF #_w5 THEN
       #Activate := FALSE;
       #Read := FALSE;
   END_IF;
   IF #_w6 AND (99 = #"Step") THEN
       #Done := FALSE;
       #Error := TRUE;
   END_IF;
   #_w7 := #_w6 AND (99 = #"Step");
   IF #_w7 THEN
       #"Step" := 0;
       #Activate := FALSE;
       #Read := FALSE;
   END_IF;
END_REGION
END_FUNCTION_BLOCK

FUNCTION_BLOCK "SAI_IND_WriteAdjustSettings"   // FB51, LAD
{ S7_Optimized_Access := 'FALSE' }
VERSION : 0.1
// stored: AutoNumber true, IsIECCheckEnabled false, SetENOAutomatically false, UDAEnableTagReadback false
   VAR_INPUT
      ID : HW_IO;   // The Profinet Device Hardware Identifier under device properties
      ScaleCapacity : Real;   // Scale capacity to be written into the transmitter
      Increment : Real;   // Increment value to be written into the transmitter
   END_VAR
   VAR_OUTPUT
      Done : Bool;   // Write process done successfully
      Error : Bool;   // Error during writing process
   END_VAR
   VAR_IN_OUT
      Write : Bool;   // Switch this bit ON to start writing
   END_VAR
   VAR DB_SPECIFIC
      Static01 : Bool;
      "Step" : Int;
   END_VAR
   VAR
      WRREC_CAP { S7_SetPoint := 'True'} : WRREC;
   END_VAR
   VAR DB_SPECIFIC
      CAP_RECORD : Real;
      INC_RECORD : Real;
      Activate : Bool;
   END_VAR
   VAR_TEMP   // added for the SCL form of the ladder/FBD networks
      _w1 : Bool;
      _w2 : Bool;
      _w3 : Bool;
      _w4 : Bool;
      _w5 : Bool;
      _w6 : Bool;
      _w7 : Bool;
   END_VAR
BEGIN

REGION Network 1: Initialization and Checking
   // Initializes FB output bits:
   // Process;
   // Error;
   // Done;
   // Check validity of scale capacity and increment values before proceeding to next step
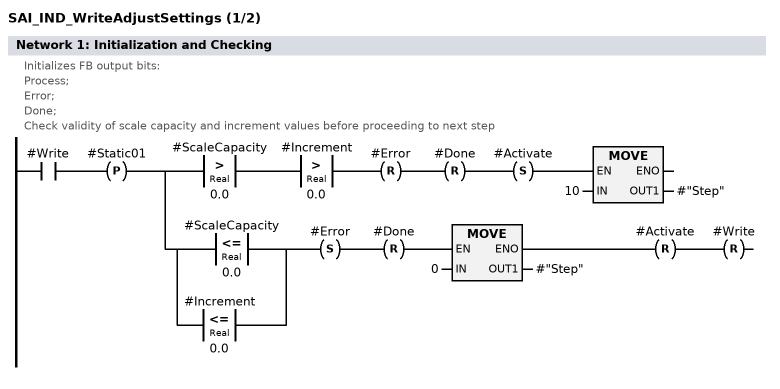
   RUNG wire#powerrail
      Contact( #Write )
      P_Trig( #Static01 )
      wire#w1
      { S7_Templates := "SrcType := Real" } GT_Contact(in1 := #ScaleCapacity, in2 := 0.0)
      { S7_Templates := "SrcType := Real" } GT_Contact(in1 := #Increment, in2 := 0.0)
      R_Coil( #Error )
      R_Coil( #Done )
      S_Coil( #Activate )
      { S7_GenerateENO := "TRUE" } Move(in := 10, out1 => #"Step")
   END_RUNG
   RUNG wire#w1
      { S7_Templates := "SrcType := Real" } LE_Contact(in1 := #ScaleCapacity, in2 := 0.0)
      wire#w2
      S_Coil( #Error )
      R_Coil( #Done )
      { S7_GenerateENO := "TRUE" } Move(in := 0, out1 => #"Step")
      R_Coil( #Activate )
      R_Coil( #Write )
   END_RUNG
   RUNG wire#w1
      { S7_Templates := "SrcType := Real" } LE_Contact(in1 := #Increment, in2 := 0.0)
   END_RUNG wire#w2
   // the same network as SCL:
   // ENO of a box is taken as its EN; it also drops when the box reports an error
   #_w1 := #Write AND NOT #Static01;   // rising edge
   #Static01 := #Write;
   IF #_w1 AND (#ScaleCapacity > 0.0) AND (#Increment > 0.0) THEN
       #Error := FALSE;
       #Done := FALSE;
       #Activate := TRUE;
       #"Step" := 10;
   END_IF;
   IF #_w1 AND ((#ScaleCapacity <= 0.0) OR (#Increment <= 0.0)) THEN
       #Error := TRUE;
       #Done := FALSE;
       #"Step" := 0;
       #Activate := FALSE;
       #Write := FALSE;
   END_IF;
END_REGION

REGION Network 2: Sequence
   // Sequence steps:
   // 10: Write in scale capacity (REAL; Index= 16#4367)
   // 20: Write in scale increment (REAL; Index= 16#4366)
   // 30: Completed the write process, DONE bit is set to TRUE
   // 99: ERROR bit is set to TRUE due to error
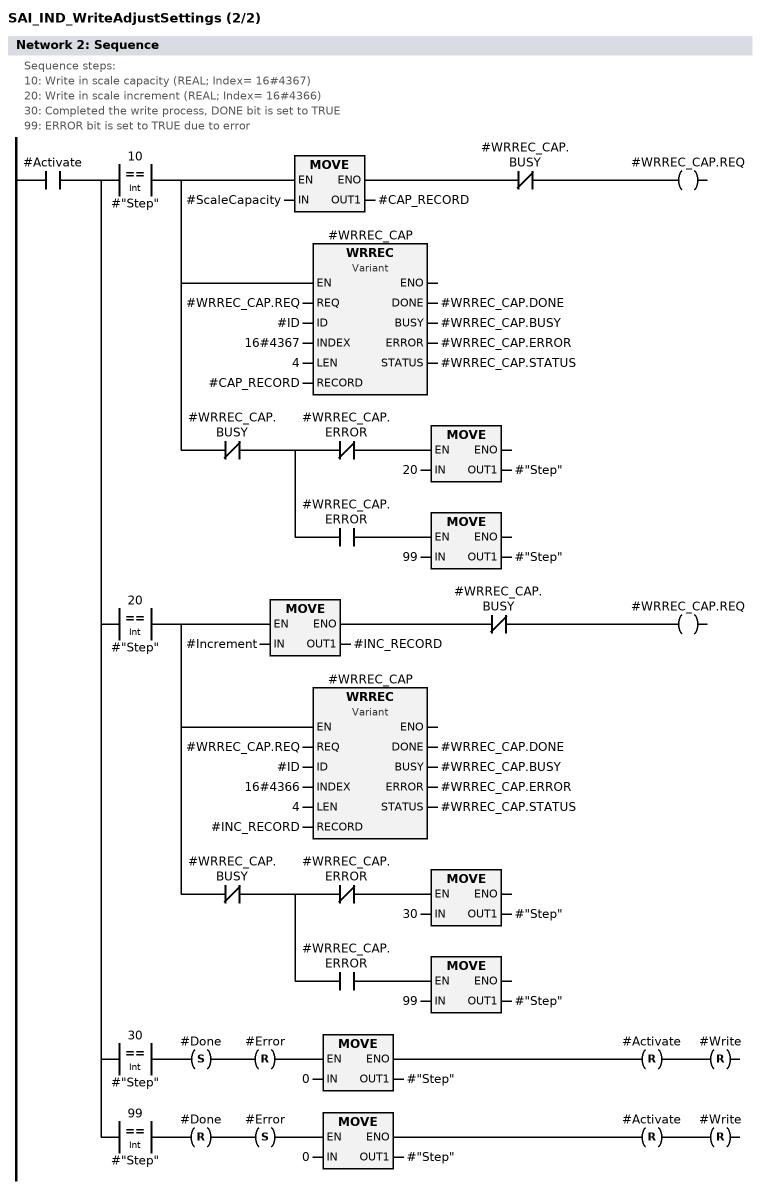
   RUNG wire#powerrail
      Contact( #Activate )
      wire#w1
      { S7_Templates := "SrcType := Int" } EQ_Contact(in1 := 10, in2 := #"Step")
      wire#w2
      { S7_GenerateENO := "TRUE" } Move(in := #ScaleCapacity, out1 => #CAP_RECORD)
      I_Contact( #WRREC_CAP.BUSY )
      Coil( #WRREC_CAP.REQ )
   END_RUNG
   RUNG wire#w2
      { S7_Templates := "[ptr_type := Variant, id_type := HW_IO, index_type := DInt, len_type := UInt]" } #WRREC_CAP.WRREC(REQ := #WRREC_CAP.REQ, ID := #ID, INDEX := 16#4367, LEN := 4, RECORD := #CAP_RECORD, DONE => #WRREC_CAP.DONE, BUSY => #WRREC_CAP.BUSY, ERROR => #WRREC_CAP.ERROR, STATUS => #WRREC_CAP.STATUS)
   END_RUNG
   RUNG wire#w2
      I_Contact( #WRREC_CAP.BUSY )
      wire#w3
      I_Contact( #WRREC_CAP.ERROR )
      { S7_GenerateENO := "TRUE" } Move(in := 20, out1 => #"Step")
   END_RUNG
   RUNG wire#w3
      Contact( #WRREC_CAP.ERROR )
      { S7_GenerateENO := "TRUE" } Move(in := 99, out1 => #"Step")
   END_RUNG
   RUNG wire#w1
      { S7_Templates := "SrcType := Int" } EQ_Contact(in1 := 20, in2 := #"Step")
      wire#w4
      { S7_GenerateENO := "TRUE" } Move(in := #Increment, out1 => #INC_RECORD)
      I_Contact( #WRREC_CAP.BUSY )
      Coil( #WRREC_CAP.REQ )
   END_RUNG
   RUNG wire#w4
      { S7_Templates := "[ptr_type := Variant, id_type := HW_IO, index_type := DInt, len_type := UInt]" } #WRREC_CAP.WRREC(REQ := #WRREC_CAP.REQ, ID := #ID, INDEX := 16#4366, LEN := 4, RECORD := #INC_RECORD, DONE => #WRREC_CAP.DONE, BUSY => #WRREC_CAP.BUSY, ERROR => #WRREC_CAP.ERROR, STATUS => #WRREC_CAP.STATUS)
   END_RUNG
   RUNG wire#w4
      I_Contact( #WRREC_CAP.BUSY )
      wire#w5
      I_Contact( #WRREC_CAP.ERROR )
      { S7_GenerateENO := "TRUE" } Move(in := 30, out1 => #"Step")
   END_RUNG
   RUNG wire#w5
      Contact( #WRREC_CAP.ERROR )
      { S7_GenerateENO := "TRUE" } Move(in := 99, out1 => #"Step")
   END_RUNG
   RUNG wire#w1
      { S7_Templates := "SrcType := Int" } EQ_Contact(in1 := 30, in2 := #"Step")
      S_Coil( #Done )
      R_Coil( #Error )
      { S7_GenerateENO := "TRUE" } Move(in := 0, out1 => #"Step")
      R_Coil( #Activate )
      R_Coil( #Write )
   END_RUNG
   RUNG wire#w1
      { S7_Templates := "SrcType := Int" } EQ_Contact(in1 := 99, in2 := #"Step")
      R_Coil( #Done )
      S_Coil( #Error )
      { S7_GenerateENO := "TRUE" } Move(in := 0, out1 => #"Step")
      R_Coil( #Activate )
      R_Coil( #Write )
   END_RUNG
   // the same network as SCL:
   // ENO of a box is taken as its EN; it also drops when the box reports an error
   #_w1 := #Activate AND (10 = #"Step");
   IF #_w1 THEN #CAP_RECORD := #ScaleCapacity; END_IF;
   #WRREC_CAP.REQ := #_w1 AND NOT #WRREC_CAP.BUSY;
   IF #_w1 THEN
       #WRREC_CAP(REQ := #WRREC_CAP.REQ,   // WRREC
                  ID := #ID,
                  INDEX := 16#4367,
                  LEN := 4,
                  RECORD := #CAP_RECORD,
                  DONE => #WRREC_CAP.DONE,
                  BUSY => #WRREC_CAP.BUSY,
                  ERROR => #WRREC_CAP.ERROR,
                  STATUS => #WRREC_CAP.STATUS);
   END_IF;
   #_w2 := #_w1 AND NOT #WRREC_CAP.BUSY;
   IF #_w2 AND NOT #WRREC_CAP.ERROR THEN #"Step" := 20; END_IF;
   IF #_w2 AND #WRREC_CAP.ERROR THEN #"Step" := 99; END_IF;
   #_w3 := #Activate AND (20 = #"Step");
   IF #_w3 THEN #INC_RECORD := #Increment; END_IF;
   #WRREC_CAP.REQ := #_w3 AND NOT #WRREC_CAP.BUSY;
   IF #_w3 THEN
       #WRREC_CAP(REQ := #WRREC_CAP.REQ,   // WRREC
                  ID := #ID,
                  INDEX := 16#4366,
                  LEN := 4,
                  RECORD := #INC_RECORD,
                  DONE => #WRREC_CAP.DONE,
                  BUSY => #WRREC_CAP.BUSY,
                  ERROR => #WRREC_CAP.ERROR,
                  STATUS => #WRREC_CAP.STATUS);
   END_IF;
   #_w4 := #_w3 AND NOT #WRREC_CAP.BUSY;
   IF #_w4 AND NOT #WRREC_CAP.ERROR THEN #"Step" := 30; END_IF;
   IF #_w4 AND #WRREC_CAP.ERROR THEN #"Step" := 99; END_IF;
   IF #Activate AND (30 = #"Step") THEN
       #Done := TRUE;
       #Error := FALSE;
   END_IF;
   #_w5 := #Activate AND (30 = #"Step");
   IF #_w5 THEN #"Step" := 0; END_IF;
   #_w6 := #Activate;
   IF #_w5 THEN
       #Activate := FALSE;
       #Write := FALSE;
   END_IF;
   IF #_w6 AND (99 = #"Step") THEN
       #Done := FALSE;
       #Error := TRUE;
   END_IF;
   #_w7 := #_w6 AND (99 = #"Step");
   IF #_w7 THEN
       #"Step" := 0;
       #Activate := FALSE;
       #Write := FALSE;
   END_IF;
END_REGION
END_FUNCTION_BLOCK

FUNCTION_BLOCK "SAI_IND_ZeroAdjust"   // FB52, LAD
TITLE = Zero Adjustment
{ S7_Optimized_Access := 'FALSE' }
VERSION : 0.1
// stored: AutoNumber true, IsIECCheckEnabled false, SetENOAutomatically false, UDAEnableTagReadback false
   VAR_INPUT
      ID : HW_IO;   // The Profinet Device Hardware Identifier under device properties
   END_VAR
   VAR_OUTPUT
      Process : Bool;   // Adjustment is in process
      Done : Bool;   // Adjustment completed successfully
      Error : Bool;
   END_VAR
   VAR_IN_OUT
      Start : Bool;   // Switch ON to start adjustment
   END_VAR
   VAR DB_SPECIFIC
      Activate : Bool;
      Status_RECORD : Int;
      Zero_RECORD : Int;
   END_VAR
   VAR
      WRREC_Zero { S7_SetPoint := 'True'} : WRREC;
      RDREC_Status { S7_SetPoint := 'True'} : RDREC;
   END_VAR
   VAR DB_SPECIFIC
      AdjustStep : SInt;
      Static01 : Bool;
      Static02 : Bool;
      Static03 : Bool;
   END_VAR
   VAR_TEMP   // added for the SCL form of the ladder/FBD networks
      _w1 : Bool;
      _w2 : Bool;
      _w3 : Bool;
      _w4 : Bool;
   END_VAR
BEGIN

REGION Network 1: Initialization
   // Initializes DONE and ERROR bits
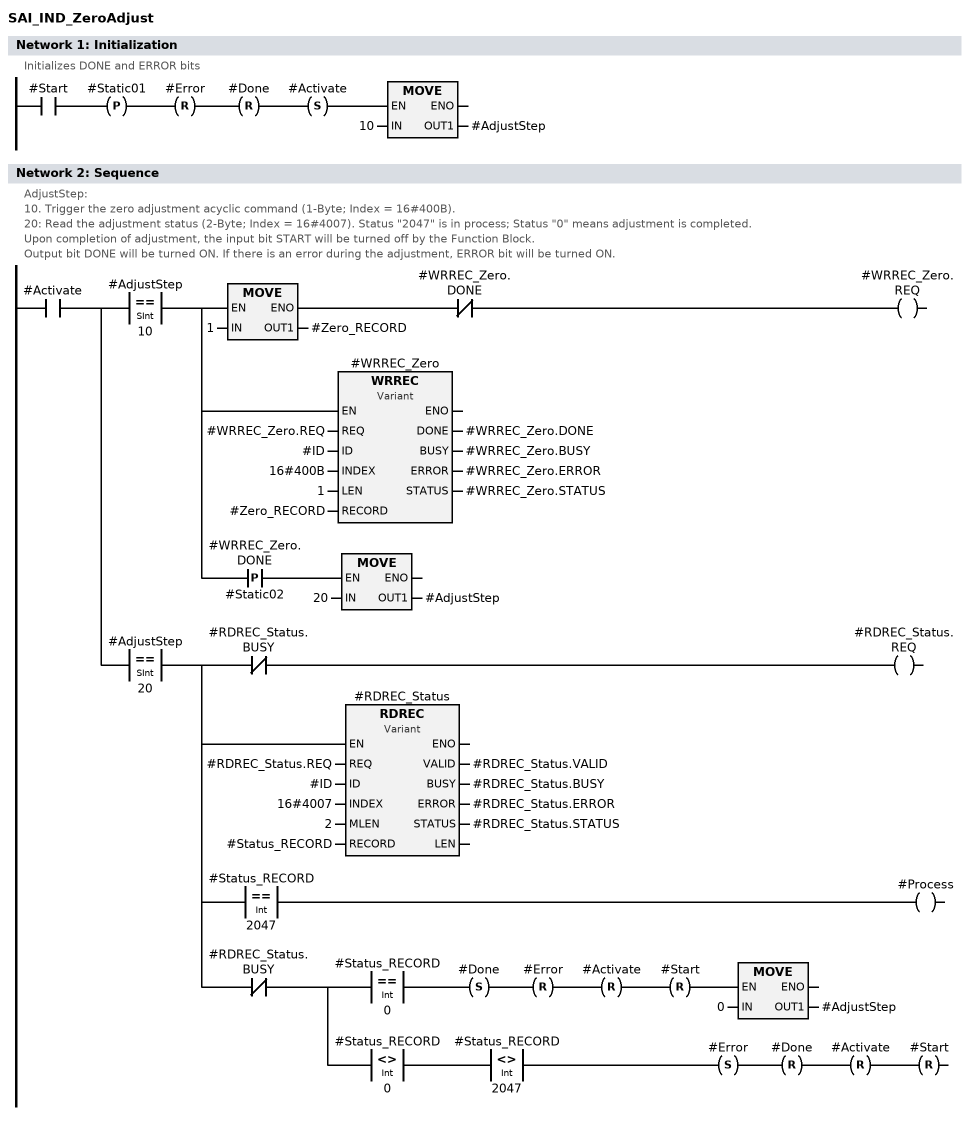
   RUNG wire#powerrail
      Contact( #Start )
      P_Trig( #Static01 )
      R_Coil( #Error )
      R_Coil( #Done )
      S_Coil( #Activate )
      { S7_GenerateENO := "TRUE" } Move(in := 10, out1 => #AdjustStep)
   END_RUNG
   // the same network as SCL:
   #_w1 := #Start AND NOT #Static01;   // rising edge
   #Static01 := #Start;
   IF #_w1 THEN
       #Error := FALSE;
       #Done := FALSE;
       #Activate := TRUE;
       #AdjustStep := 10;
   END_IF;
END_REGION

REGION Network 2: Sequence
   // AdjustStep:
   // 
   // 10. Trigger the zero adjustment acyclic command (1-Byte; Index = 16#400B). 
   // 
   // 20: Read the adjustment status (2-Byte; Index = 16#4007). Status "2047" is in process; Status "0" means adjustment is completed.
   // Upon completion of adjustment, the input bit START will be turned off by the Function Block.
   // Output bit DONE will be turned ON. If there is an error during the adjustment, ERROR bit will be turned ON.
   RUNG wire#powerrail
      Contact( #Activate )
      wire#w1
      { S7_Templates := "SrcType := SInt" } EQ_Contact(in1 := #AdjustStep, in2 := 10)
      wire#w2
      Move(in := 1, out1 => #Zero_RECORD)
      I_Contact( #WRREC_Zero.DONE )
      Coil( #WRREC_Zero.REQ )
   END_RUNG
   RUNG wire#w2
      { S7_Templates := "[ptr_type := Variant, id_type := HW_IO, index_type := DInt, len_type := UInt]" } #WRREC_Zero.WRREC(REQ := #WRREC_Zero.REQ, ID := #ID, INDEX := 16#400B, LEN := 1, RECORD := #Zero_RECORD, DONE => #WRREC_Zero.DONE, BUSY => #WRREC_Zero.BUSY, ERROR => #WRREC_Zero.ERROR, STATUS => #WRREC_Zero.STATUS)
   END_RUNG
   RUNG wire#w2
      P_Contact(operand := #WRREC_Zero.DONE, bit := #Static02)
      Move(in := 20, out1 => #AdjustStep)
   END_RUNG
   RUNG wire#w1
      { S7_Templates := "SrcType := SInt" } EQ_Contact(in1 := #AdjustStep, in2 := 20)
      wire#w3
      I_Contact( #RDREC_Status.BUSY )
      Coil( #RDREC_Status.REQ )
   END_RUNG
   RUNG wire#w3
      { S7_Templates := "[ptr_type := Variant, id_type := HW_IO, index_type := DInt, len_type := UInt]" } #RDREC_Status.RDREC(REQ := #RDREC_Status.REQ, ID := #ID, INDEX := 16#4007, MLEN := 2, RECORD := #Status_RECORD, VALID => #RDREC_Status.VALID, BUSY => #RDREC_Status.BUSY, ERROR => #RDREC_Status.ERROR, STATUS => #RDREC_Status.STATUS, LEN =>)
   END_RUNG
   RUNG wire#w3
      { S7_Templates := "SrcType := Int" } EQ_Contact(in1 := #Status_RECORD, in2 := 2047)
      Coil( #Process )
   END_RUNG
   RUNG wire#w3
      I_Contact( #RDREC_Status.BUSY )
      wire#w4
      { S7_Templates := "SrcType := Int" } EQ_Contact(in1 := #Status_RECORD, in2 := 0)
      S_Coil( #Done )
      R_Coil( #Error )
      R_Coil( #Activate )
      R_Coil( #Start )
      Move(in := 0, out1 => #AdjustStep)
   END_RUNG
   RUNG wire#w4
      { S7_Templates := "SrcType := Int" } NE_Contact(in1 := #Status_RECORD, in2 := 0)
      { S7_Templates := "SrcType := Int" } NE_Contact(in1 := #Status_RECORD, in2 := 2047)
      S_Coil( #Error )
      R_Coil( #Done )
      R_Coil( #Activate )
      R_Coil( #Start )
   END_RUNG
   // the same network as SCL:
   #_w1 := #Activate AND (#AdjustStep = 10);
   IF #_w1 THEN #Zero_RECORD := 1; END_IF;
   #WRREC_Zero.REQ := #_w1 AND NOT #WRREC_Zero.DONE;
   IF #_w1 THEN
       #WRREC_Zero(REQ := #WRREC_Zero.REQ,   // WRREC
                   ID := #ID,
                   INDEX := 16#400B,
                   LEN := 1,
                   RECORD := #Zero_RECORD,
                   DONE => #WRREC_Zero.DONE,
                   BUSY => #WRREC_Zero.BUSY,
                   ERROR => #WRREC_Zero.ERROR,
                   STATUS => #WRREC_Zero.STATUS);
   END_IF;
   #_w2 := #_w1 AND #WRREC_Zero.DONE AND NOT #Static02;   // rising edge of #WRREC_Zero.DONE
   #Static02 := #WRREC_Zero.DONE;
   IF #_w2 THEN #AdjustStep := 20; END_IF;
   #_w3 := #Activate AND (#AdjustStep = 20);
   #RDREC_Status.REQ := #_w3 AND NOT #RDREC_Status.BUSY;
   IF #_w3 THEN
       #RDREC_Status(REQ := #RDREC_Status.REQ,   // RDREC
                     ID := #ID,
                     INDEX := 16#4007,
                     MLEN := 2,
                     RECORD := #Status_RECORD,
                     VALID => #RDREC_Status.VALID,
                     BUSY => #RDREC_Status.BUSY,
                     ERROR => #RDREC_Status.ERROR,
                     STATUS => #RDREC_Status.STATUS);
   END_IF;
   #Process := #_w3 AND (#Status_RECORD = 2047);
   #_w4 := #_w3 AND NOT #RDREC_Status.BUSY;
   IF #_w4 AND (#Status_RECORD = 0) THEN
       #Done := TRUE;
       #Error := FALSE;
       #Activate := FALSE;
       #Start := FALSE;
       #AdjustStep := 0;
   END_IF;
   IF #_w4 AND (#Status_RECORD <> 0) AND (#Status_RECORD <> 2047) THEN
       #Error := TRUE;
       #Done := FALSE;
       #Activate := FALSE;
       #Start := FALSE;
   END_IF;
END_REGION
END_FUNCTION_BLOCK

FUNCTION_BLOCK "SAI_IND_SpanAdjust"   // FB55, LAD
TITLE = Span and Linearity Adjustment (Multi-Point Selectable)
{ S7_Optimized_Access := 'FALSE' }
VERSION : 0.1
// stored: AutoNumber true, IsIECCheckEnabled false, SetENOAutomatically false, UDAEnableTagReadback false
   VAR_INPUT
      ID : HW_IO;   // The Profinet Device Hardware Identifier under device properties
      Hi_Weight : Real;   // The highest adjustment weight, or the Span value
      Mid_Weight : Real;   // The 4th adjustment weight
      Low_Weight : Real;   // The 3rd adjustment weight
      xLow_Weight : Real;   // The 2nd adjustment weight
   END_VAR
   VAR_OUTPUT
      CurrentPoint : Int;   // Current point to be adjusted (Minimum 2 points; maximum 5 points; zero point is the 1st point)
      CurrentWeight : Real;   // Current adjustment weight to be loaded onto the scale
      LoadWeight : Bool;   // Load the next adjustment weight according to value shown in CurrentWeight
      Process : Bool;   // Weight Transmitter is performing adjustment
      Done : Bool;   // Linearity Adjustment has been completed successfully
      Error : Bool;   // Adjustment can not proceed due to incomplete input parameters, check LinearityRange and all the adjustment weight values
      Cancelled : Bool;   // Adjustment process has been cancelled successfully
   END_VAR
   VAR_IN_OUT
      LinearityRange : Int;   // Number of linearity points to be adjusted: 0:none, 1:3 point, 2:4 point, 3:5 point
      Start : Bool;   // Trigger this bit ON to start performing linearity adjustment; this bit will be turned off automatically after completion
      ConfirmWeight : Bool;   // Switch ON this bit as an acknowledgement that new adjustment weight has being loaded
      Cancel : Bool;   // Cancel/ Abort adjustment process, toggle ON
   END_VAR
   VAR DB_SPECIFIC
      Activate : Bool;
   END_VAR
   VAR
      WRREC_SpanAdjust { S7_SetPoint := 'True'} : WRREC;
      RDREC_Status { S7_SetPoint := 'True'} : RDREC;
   END_VAR
   VAR DB_SPECIFIC
      IEC_Timer_1_Instance { S7_SetPoint := 'True'} : IEC_TIMER;
      AdjustStep : SInt;
      Static01 : Bool;
      Static02 : Bool;
      Static03 : Bool;
      Static04 : Bool;
      Static05 : Bool;
      Static06 : Bool;
      Static07 : Bool;
      Static08 : Bool;
      Validate_REC : SInt;
      Abort_REC : SInt;
      Check01 : Bool;
      Check02 : Bool;
      AdjustmentStatus : Int;
      CurrentPoint_0 : Int;
      CurrentWeight_0 : Real;
   END_VAR
   VAR_TEMP   // added for the SCL form of the ladder/FBD networks
      _w1 : Bool;
      _w2 : Bool;
      _w3 : Bool;
      _w4 : Bool;
      _w5 : Bool;
      _w6 : Bool;
      _w7 : Bool;
      _w8 : Bool;
      _w9 : Bool;
      _w10 : Bool;
      _w11 : Bool;
      _w12 : Bool;
      _w13 : Bool;
   END_VAR
BEGIN

REGION Network 1: Initialization
   // Initializes FB output bits:
   // Process;
   // Error;
   // Done;
   // Cancelled
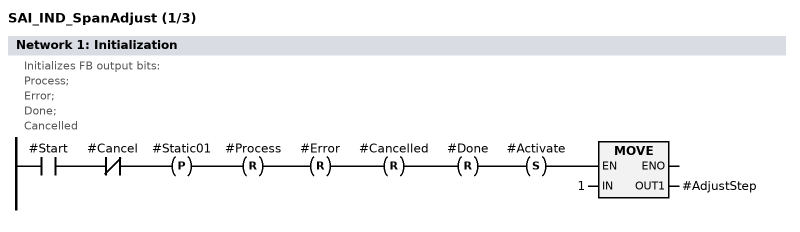
   RUNG wire#powerrail
      Contact( #Start )
      I_Contact( #Cancel )
      P_Trig( #Static01 )
      R_Coil( #Process )
      R_Coil( #Error )
      R_Coil( #Cancelled )
      R_Coil( #Done )
      S_Coil( #Activate )
      { S7_GenerateENO := "TRUE" } Move(in := 1, out1 => #AdjustStep)
   END_RUNG
   // the same network as SCL:
   #_w1 := #Start AND NOT #Cancel;
   #_w2 := #_w1 AND NOT #Static01;   // rising edge
   #Static01 := #_w1;
   IF #_w2 THEN
       #Process := FALSE;
       #Error := FALSE;
       #Cancelled := FALSE;
       #Done := FALSE;
       #Activate := TRUE;
       #AdjustStep := 1;
   END_IF;
END_REGION

REGION Network 2: Sequence
   // AdjustStep = 1: Check all the input parameters for LinearityRange and adjustment weights (Hi_Weight, Mid_Weight, Low_Weight, xLow_Weight)
   // AdjustStep = 2: Initializes all the control bits
   // AdjustStep = 3: Write in the LinearityRange into the transmitter (2-byte; Index: 16#400A)
   // AdjustStep = 4: Updates the CurrentPoint and CurrentWeight (new reference weight) and wait for user to trigger ConfirmWeight input bit
   // AdjustStep = 5: Start the adjustment process according to the CurrentWeight (REAL; Index: 16#4009)
   // AdjustStep = 6: After adjusted all the required reference weights, validate the adjustment (2-byte; Index: 16#4010)
   // AdjustStep = 7: Adjustment is completed successfully, set DONE bit to TRUE
   // AdjustStep = 8; Adjustment failed with error, set ERROR bit to TRUE
   // AdjustStep >= 4: Reading the adjustment status continuously (2-byte; Index: 16#4007)
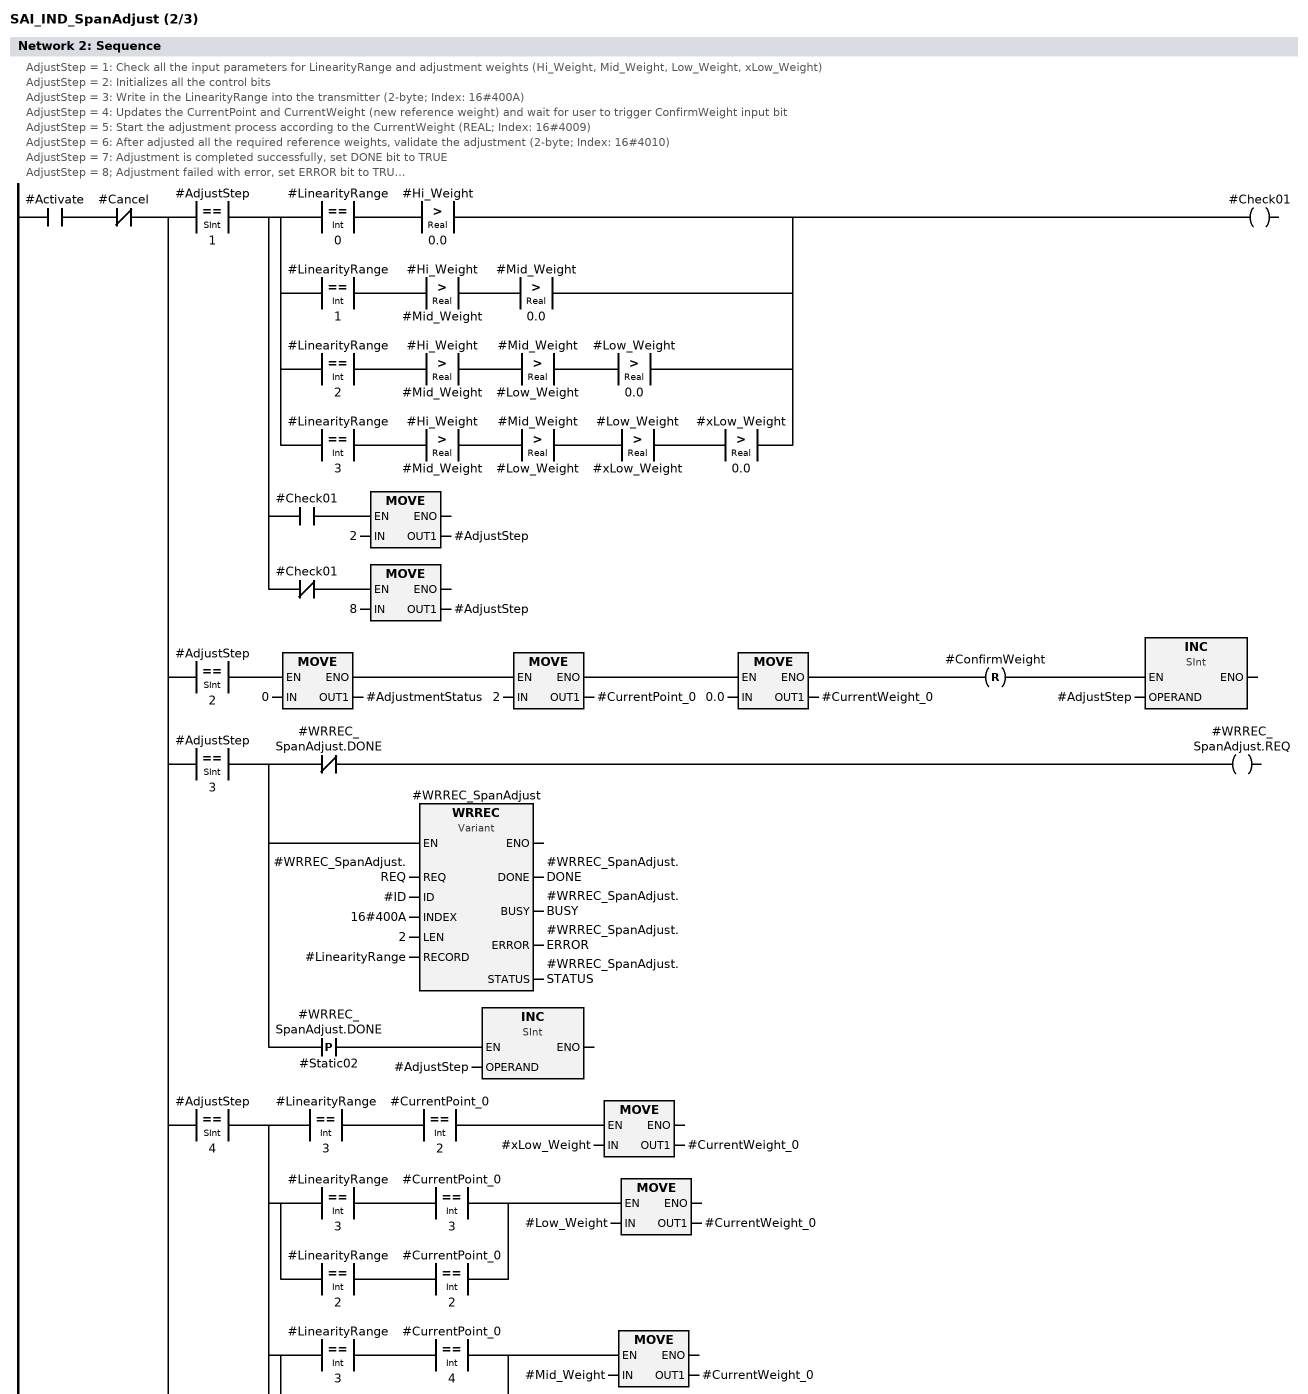
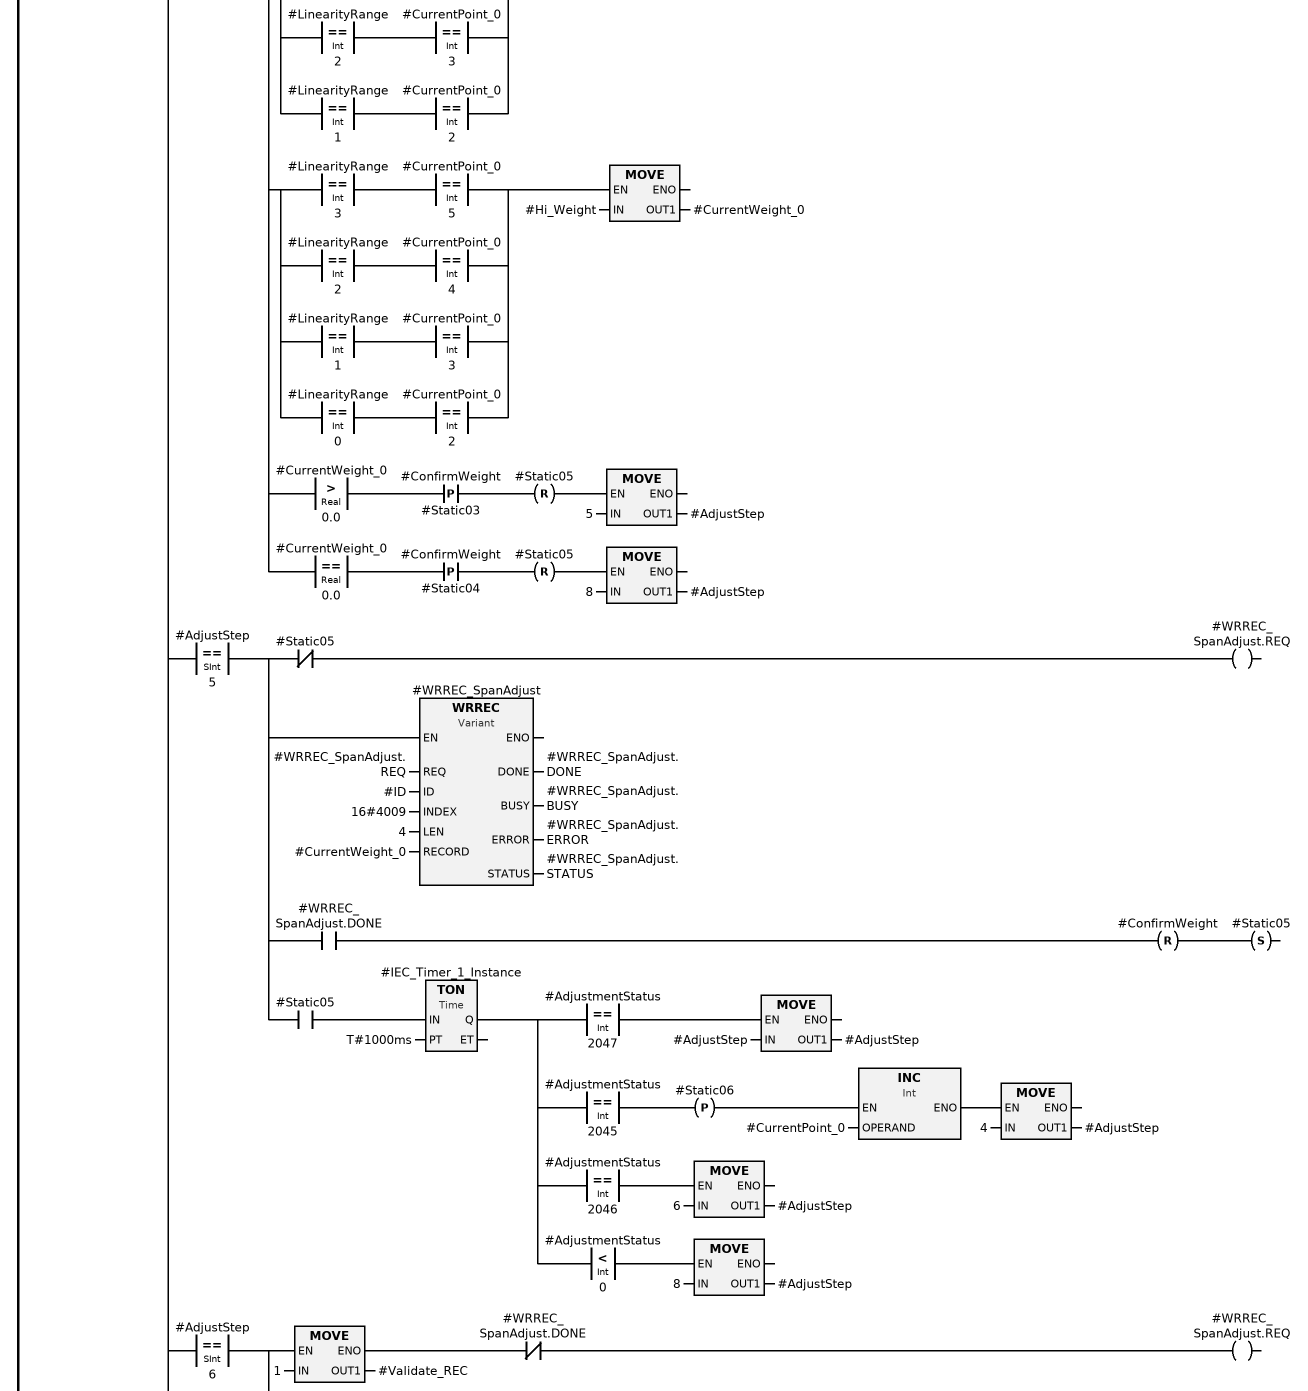
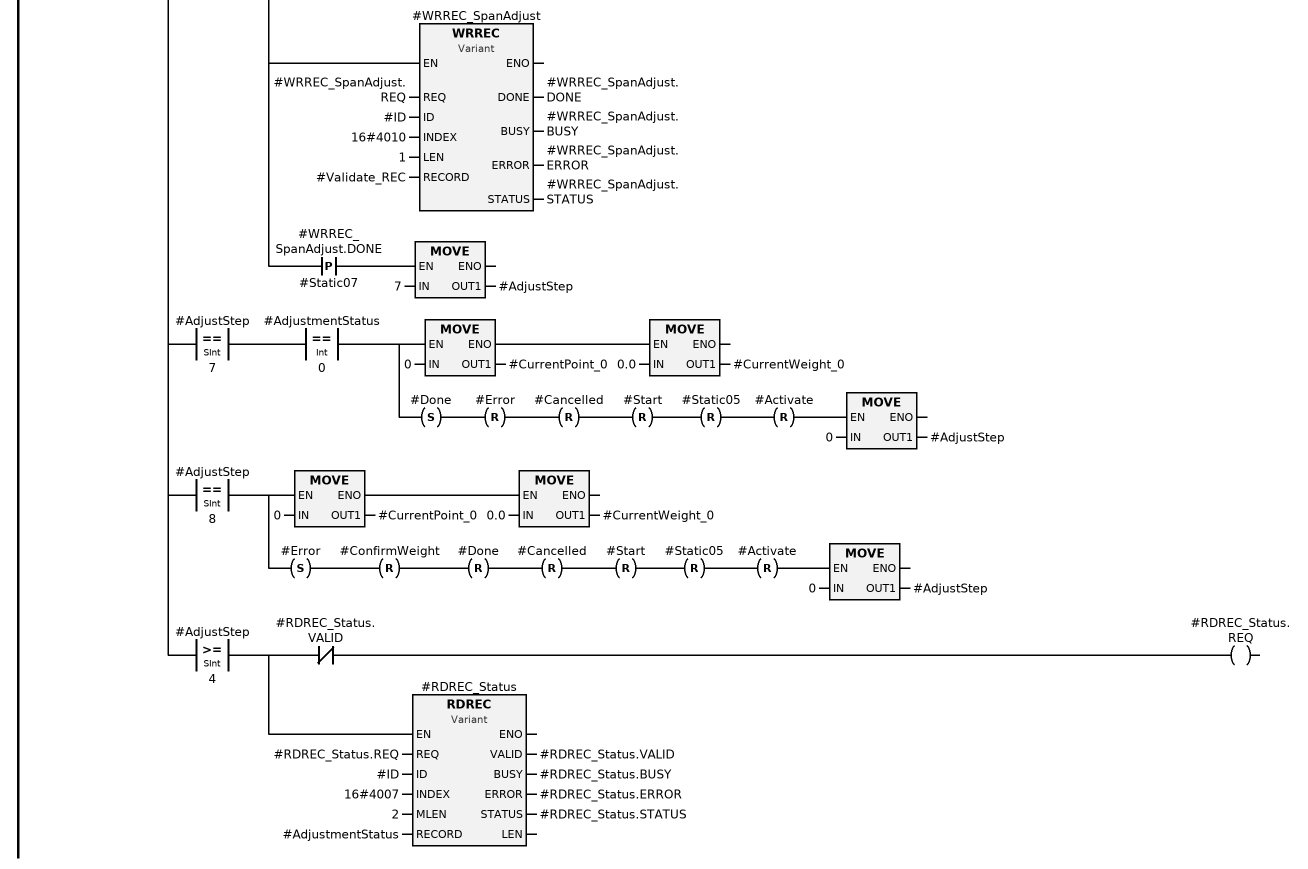
   RUNG wire#powerrail
      Contact( #Activate )
      I_Contact( #Cancel )
      wire#w1
      { S7_Templates := "SrcType := SInt" } EQ_Contact(in1 := #AdjustStep, in2 := 1)
      wire#w2
      { S7_Templates := "SrcType := Int" } EQ_Contact(in1 := #LinearityRange, in2 := 0)
      { S7_Templates := "SrcType := Real" } GT_Contact(in1 := #Hi_Weight, in2 := 0.0)
      wire#w3
      Coil( #Check01 )
   END_RUNG
   RUNG wire#w2
      { S7_Templates := "SrcType := Int" } EQ_Contact(in1 := #LinearityRange, in2 := 1)
      { S7_Templates := "SrcType := Real" } GT_Contact(in1 := #Hi_Weight, in2 := #Mid_Weight)
      { S7_Templates := "SrcType := Real" } GT_Contact(in1 := #Mid_Weight, in2 := 0.0)
   END_RUNG wire#w3
   RUNG wire#w2
      { S7_Templates := "SrcType := Int" } EQ_Contact(in1 := #LinearityRange, in2 := 2)
      { S7_Templates := "SrcType := Real" } GT_Contact(in1 := #Hi_Weight, in2 := #Mid_Weight)
      { S7_Templates := "SrcType := Real" } GT_Contact(in1 := #Mid_Weight, in2 := #Low_Weight)
      { S7_Templates := "SrcType := Real" } GT_Contact(in1 := #Low_Weight, in2 := 0.0)
   END_RUNG wire#w3
   RUNG wire#w2
      { S7_Templates := "SrcType := Int" } EQ_Contact(in1 := #LinearityRange, in2 := 3)
      { S7_Templates := "SrcType := Real" } GT_Contact(in1 := #Hi_Weight, in2 := #Mid_Weight)
      { S7_Templates := "SrcType := Real" } GT_Contact(in1 := #Mid_Weight, in2 := #Low_Weight)
      { S7_Templates := "SrcType := Real" } GT_Contact(in1 := #Low_Weight, in2 := #xLow_Weight)
      { S7_Templates := "SrcType := Real" } GT_Contact(in1 := #xLow_Weight, in2 := 0.0)
   END_RUNG wire#w3
   RUNG wire#w2
      Contact( #Check01 )
      Move(in := 2, out1 => #AdjustStep)
   END_RUNG
   RUNG wire#w2
      I_Contact( #Check01 )
      Move(in := 8, out1 => #AdjustStep)
   END_RUNG
   RUNG wire#w1
      { S7_Templates := "SrcType := SInt" } EQ_Contact(in1 := #AdjustStep, in2 := 2)
      Move(in := 0, out1 => #AdjustmentStatus)
      Move(in := 2, out1 => #CurrentPoint_0)
      Move(in := 0.0, out1 => #CurrentWeight_0)
      R_Coil( #ConfirmWeight )
      { S7_Templates := "DestType := SInt" } Inc( #AdjustStep )
   END_RUNG
   RUNG wire#w1
      { S7_Templates := "SrcType := SInt" } EQ_Contact(in1 := #AdjustStep, in2 := 3)
      wire#w4
      I_Contact( #WRREC_SpanAdjust.DONE )
      Coil( #WRREC_SpanAdjust.REQ )
   END_RUNG
   RUNG wire#w4
      { S7_Templates := "[ptr_type := Variant, id_type := HW_IO, index_type := DInt, len_type := UInt]" } #WRREC_SpanAdjust.WRREC(REQ := #WRREC_SpanAdjust.REQ, ID := #ID, INDEX := 16#400A, LEN := 2, RECORD := #LinearityRange, DONE => #WRREC_SpanAdjust.DONE, BUSY => #WRREC_SpanAdjust.BUSY, ERROR => #WRREC_SpanAdjust.ERROR, STATUS => #WRREC_SpanAdjust.STATUS)
   END_RUNG
   RUNG wire#w4
      P_Contact(operand := #WRREC_SpanAdjust.DONE, bit := #Static02)
      { S7_Templates := "DestType := SInt" } Inc( #AdjustStep )
   END_RUNG
   RUNG wire#w1
      { S7_Templates := "SrcType := SInt" } EQ_Contact(in1 := #AdjustStep, in2 := 4)
      wire#w5
      { S7_Templates := "SrcType := Int" } EQ_Contact(in1 := #LinearityRange, in2 := 3)
      { S7_Templates := "SrcType := Int" } EQ_Contact(in1 := #CurrentPoint_0, in2 := 2)
      Move(in := #xLow_Weight, out1 => #CurrentWeight_0)
   END_RUNG
   RUNG wire#w5
      { S7_Templates := "SrcType := Int" } EQ_Contact(in1 := #LinearityRange, in2 := 3)
      { S7_Templates := "SrcType := Int" } EQ_Contact(in1 := #CurrentPoint_0, in2 := 3)
      wire#w6
      Move(in := #Low_Weight, out1 => #CurrentWeight_0)
   END_RUNG
   RUNG wire#w5
      { S7_Templates := "SrcType := Int" } EQ_Contact(in1 := #LinearityRange, in2 := 2)
      { S7_Templates := "SrcType := Int" } EQ_Contact(in1 := #CurrentPoint_0, in2 := 2)
   END_RUNG wire#w6
   RUNG wire#w5
      { S7_Templates := "SrcType := Int" } EQ_Contact(in1 := #LinearityRange, in2 := 3)
      { S7_Templates := "SrcType := Int" } EQ_Contact(in1 := #CurrentPoint_0, in2 := 4)
      wire#w7
      Move(in := #Mid_Weight, out1 => #CurrentWeight_0)
   END_RUNG
   RUNG wire#w5
      { S7_Templates := "SrcType := Int" } EQ_Contact(in1 := #LinearityRange, in2 := 2)
      { S7_Templates := "SrcType := Int" } EQ_Contact(in1 := #CurrentPoint_0, in2 := 3)
   END_RUNG wire#w7
   RUNG wire#w5
      { S7_Templates := "SrcType := Int" } EQ_Contact(in1 := #LinearityRange, in2 := 1)
      { S7_Templates := "SrcType := Int" } EQ_Contact(in1 := #CurrentPoint_0, in2 := 2)
   END_RUNG wire#w7
   RUNG wire#w5
      { S7_Templates := "SrcType := Int" } EQ_Contact(in1 := #LinearityRange, in2 := 3)
      { S7_Templates := "SrcType := Int" } EQ_Contact(in1 := #CurrentPoint_0, in2 := 5)
      wire#w8
      Move(in := #Hi_Weight, out1 => #CurrentWeight_0)
   END_RUNG
   RUNG wire#w5
      { S7_Templates := "SrcType := Int" } EQ_Contact(in1 := #LinearityRange, in2 := 2)
      { S7_Templates := "SrcType := Int" } EQ_Contact(in1 := #CurrentPoint_0, in2 := 4)
   END_RUNG wire#w8
   RUNG wire#w5
      { S7_Templates := "SrcType := Int" } EQ_Contact(in1 := #LinearityRange, in2 := 1)
      { S7_Templates := "SrcType := Int" } EQ_Contact(in1 := #CurrentPoint_0, in2 := 3)
   END_RUNG wire#w8
   RUNG wire#w5
      { S7_Templates := "SrcType := Int" } EQ_Contact(in1 := #LinearityRange, in2 := 0)
      { S7_Templates := "SrcType := Int" } EQ_Contact(in1 := #CurrentPoint_0, in2 := 2)
   END_RUNG wire#w8
   RUNG wire#w5
      { S7_Templates := "SrcType := Real" } GT_Contact(in1 := #CurrentWeight_0, in2 := 0.0)
      P_Contact(operand := #ConfirmWeight, bit := #Static03)
      R_Coil( #Static05 )
      Move(in := 5, out1 => #AdjustStep)
   END_RUNG
   RUNG wire#w5
      { S7_Templates := "SrcType := Real" } EQ_Contact(in1 := #CurrentWeight_0, in2 := 0.0)
      P_Contact(operand := #ConfirmWeight, bit := #Static04)
      R_Coil( #Static05 )
      Move(in := 8, out1 => #AdjustStep)
   END_RUNG
   RUNG wire#w1
      { S7_Templates := "SrcType := SInt" } EQ_Contact(in1 := #AdjustStep, in2 := 5)
      wire#w9
      I_Contact( #Static05 )
      Coil( #WRREC_SpanAdjust.REQ )
   END_RUNG
   RUNG wire#w9
      { S7_Templates := "[ptr_type := Variant, id_type := HW_IO, index_type := DInt, len_type := UInt]" } #WRREC_SpanAdjust.WRREC(REQ := #WRREC_SpanAdjust.REQ, ID := #ID, INDEX := 16#4009, LEN := 4, RECORD := #CurrentWeight_0, DONE => #WRREC_SpanAdjust.DONE, BUSY => #WRREC_SpanAdjust.BUSY, ERROR => #WRREC_SpanAdjust.ERROR, STATUS => #WRREC_SpanAdjust.STATUS)
   END_RUNG
   RUNG wire#w9
      Contact( #WRREC_SpanAdjust.DONE )
      R_Coil( #ConfirmWeight )
      S_Coil( #Static05 )
   END_RUNG
   RUNG wire#w9
      Contact( #Static05 )
      { S7_Templates := "time_type := Time" } #IEC_Timer_1_Instance.TON(pt := T#1000ms, et =>)
      wire#w10
      { S7_Templates := "SrcType := Int" } EQ_Contact(in1 := #AdjustmentStatus, in2 := 2047)
      Move(in := #AdjustStep, out1 => #AdjustStep)
   END_RUNG
   RUNG wire#w10
      { S7_Templates := "SrcType := Int" } EQ_Contact(in1 := #AdjustmentStatus, in2 := 2045)
      P_Trig( #Static06 )
      { S7_Templates := "DestType := Int" } Inc( #CurrentPoint_0 )
      Move(in := 4, out1 => #AdjustStep)
   END_RUNG
   RUNG wire#w10
      { S7_Templates := "SrcType := Int" } EQ_Contact(in1 := #AdjustmentStatus, in2 := 2046)
      Move(in := 6, out1 => #AdjustStep)
   END_RUNG
   RUNG wire#w10
      { S7_Templates := "SrcType := Int" } LT_Contact(in1 := #AdjustmentStatus, in2 := 0)
      Move(in := 8, out1 => #AdjustStep)
   END_RUNG
   RUNG wire#w1
      { S7_Templates := "SrcType := SInt" } EQ_Contact(in1 := #AdjustStep, in2 := 6)
      wire#w11
      Move(in := 1, out1 => #Validate_REC)
      I_Contact( #WRREC_SpanAdjust.DONE )
      Coil( #WRREC_SpanAdjust.REQ )
   END_RUNG
   RUNG wire#w11
      { S7_Templates := "[ptr_type := Variant, id_type := HW_IO, index_type := DInt, len_type := UInt]" } #WRREC_SpanAdjust.WRREC(REQ := #WRREC_SpanAdjust.REQ, ID := #ID, INDEX := 16#4010, LEN := 1, RECORD := #Validate_REC, DONE => #WRREC_SpanAdjust.DONE, BUSY => #WRREC_SpanAdjust.BUSY, ERROR => #WRREC_SpanAdjust.ERROR, STATUS => #WRREC_SpanAdjust.STATUS)
   END_RUNG
   RUNG wire#w11
      P_Contact(operand := #WRREC_SpanAdjust.DONE, bit := #Static07)
      Move(in := 7, out1 => #AdjustStep)
   END_RUNG
   RUNG wire#w1
      { S7_Templates := "SrcType := SInt" } EQ_Contact(in1 := #AdjustStep, in2 := 7)
      { S7_Templates := "SrcType := Int" } EQ_Contact(in1 := #AdjustmentStatus, in2 := 0)
      wire#w12
      Move(in := 0, out1 => #CurrentPoint_0)
      Move(in := 0.0, out1 => #CurrentWeight_0)
   END_RUNG
   RUNG wire#w12
      S_Coil( #Done )
      R_Coil( #Error )
      R_Coil( #Cancelled )
      R_Coil( #Start )
      R_Coil( #Static05 )
      R_Coil( #Activate )
      Move(in := 0, out1 => #AdjustStep)
   END_RUNG
   RUNG wire#w1
      { S7_Templates := "SrcType := SInt" } EQ_Contact(in1 := #AdjustStep, in2 := 8)
      wire#w13
      Move(in := 0, out1 => #CurrentPoint_0)
      Move(in := 0.0, out1 => #CurrentWeight_0)
   END_RUNG
   RUNG wire#w13
      S_Coil( #Error )
      R_Coil( #ConfirmWeight )
      R_Coil( #Done )
      R_Coil( #Cancelled )
      R_Coil( #Start )
      R_Coil( #Static05 )
      R_Coil( #Activate )
      Move(in := 0, out1 => #AdjustStep)
   END_RUNG
   RUNG wire#w1
      { S7_Templates := "SrcType := SInt" } GE_Contact(in1 := #AdjustStep, in2 := 4)
      wire#w14
      I_Contact( #RDREC_Status.VALID )
      Coil( #RDREC_Status.REQ )
   END_RUNG
   RUNG wire#w14
      { S7_Templates := "[ptr_type := Variant, id_type := HW_IO, index_type := DInt, len_type := UInt]" } #RDREC_Status.RDREC(REQ := #RDREC_Status.REQ, ID := #ID, INDEX := 16#4007, MLEN := 2, RECORD := #AdjustmentStatus, VALID => #RDREC_Status.VALID, BUSY => #RDREC_Status.BUSY, ERROR => #RDREC_Status.ERROR, STATUS => #RDREC_Status.STATUS, LEN =>)
   END_RUNG
   // the same network as SCL:
   #_w1 := #Activate AND NOT #Cancel;
   #_w2 := #_w1 AND (#AdjustStep = 1);
   #Check01 := #_w2 AND (((#LinearityRange = 0) AND (#Hi_Weight > 0.0)) OR ((#LinearityRange = 1) AND (#Hi_Weight > #Mid_Weight) AND (#Mid_Weight > 0.0)) OR ((#LinearityRange = 2) AND (#Hi_Weight > #Mid_Weight) AND (#Mid_Weight > #Low_Weight) AND (#Low_Weight > 0.0)) OR ((#LinearityRange = 3) AND (#Hi_Weight > #Mid_Weight) AND (#Mid_Weight > #Low_Weight) AND (#Low_Weight > #xLow_Weight) AND (#xLow_Weight > 0.0)));
   IF #_w2 AND #Check01 THEN #AdjustStep := 2; END_IF;
   IF #_w2 AND NOT #Check01 THEN #AdjustStep := 8; END_IF;
   IF #_w1 AND (#AdjustStep = 2) THEN
       #AdjustmentStatus := 0;
       #CurrentPoint_0 := 2;
       #CurrentWeight_0 := 0.0;
       #ConfirmWeight := FALSE;
       #AdjustStep := #AdjustStep + 1;
   END_IF;
   #_w3 := #_w1 AND (#AdjustStep = 3);
   #WRREC_SpanAdjust.REQ := #_w3 AND NOT #WRREC_SpanAdjust.DONE;
   IF #_w3 THEN
       #WRREC_SpanAdjust(REQ := #WRREC_SpanAdjust.REQ,   // WRREC
                         ID := #ID,
                         INDEX := 16#400A,
                         LEN := 2,
                         RECORD := #LinearityRange,
                         DONE => #WRREC_SpanAdjust.DONE,
                         BUSY => #WRREC_SpanAdjust.BUSY,
                         ERROR => #WRREC_SpanAdjust.ERROR,
                         STATUS => #WRREC_SpanAdjust.STATUS);
   END_IF;
   #_w4 := #_w3 AND #WRREC_SpanAdjust.DONE AND NOT #Static02;   // rising edge of #WRREC_SpanAdjust.DONE
   #Static02 := #WRREC_SpanAdjust.DONE;
   IF #_w4 THEN #AdjustStep := #AdjustStep + 1; END_IF;
   #_w5 := #_w1 AND (#AdjustStep = 4);
   IF #_w5 AND (#LinearityRange = 3) AND (#CurrentPoint_0 = 2) THEN #CurrentWeight_0 := #xLow_Weight; END_IF;
   IF #_w5 AND (((#LinearityRange = 3) AND (#CurrentPoint_0 = 3)) OR ((#LinearityRange = 2) AND (#CurrentPoint_0 = 2))) THEN
       #CurrentWeight_0 := #Low_Weight;
   END_IF;
   IF #_w5 AND (((#LinearityRange = 3) AND (#CurrentPoint_0 = 4)) OR ((#LinearityRange = 2) AND (#CurrentPoint_0 = 3)) OR ((#LinearityRange = 1) AND (#CurrentPoint_0 = 2))) THEN
       #CurrentWeight_0 := #Mid_Weight;
   END_IF;
   IF #_w5 AND (((#LinearityRange = 3) AND (#CurrentPoint_0 = 5)) OR ((#LinearityRange = 2) AND (#CurrentPoint_0 = 4)) OR ((#LinearityRange = 1) AND (#CurrentPoint_0 = 3)) OR ((#LinearityRange = 0) AND (#CurrentPoint_0 = 2))) THEN
       #CurrentWeight_0 := #Hi_Weight;
   END_IF;
   #_w6 := #_w5 AND (#CurrentWeight_0 > 0.0) AND #ConfirmWeight AND NOT #Static03;   // rising edge of #ConfirmWeight
   #Static03 := #ConfirmWeight;
   IF #_w6 THEN
       #Static05 := FALSE;
       #AdjustStep := 5;
   END_IF;
   #_w7 := #_w5 AND (#CurrentWeight_0 = 0.0) AND #ConfirmWeight AND NOT #Static04;   // rising edge of #ConfirmWeight
   #Static04 := #ConfirmWeight;
   IF #_w7 THEN
       #Static05 := FALSE;
       #AdjustStep := 8;
   END_IF;
   #_w8 := #_w1 AND (#AdjustStep = 5);
   #WRREC_SpanAdjust.REQ := #_w8 AND NOT #Static05;
   IF #_w8 THEN
       #WRREC_SpanAdjust(REQ := #WRREC_SpanAdjust.REQ,   // WRREC
                         ID := #ID,
                         INDEX := 16#4009,
                         LEN := 4,
                         RECORD := #CurrentWeight_0,
                         DONE => #WRREC_SpanAdjust.DONE,
                         BUSY => #WRREC_SpanAdjust.BUSY,
                         ERROR => #WRREC_SpanAdjust.ERROR,
                         STATUS => #WRREC_SpanAdjust.STATUS);
   END_IF;
   IF #_w8 AND #WRREC_SpanAdjust.DONE THEN
       #ConfirmWeight := FALSE;
       #Static05 := TRUE;
   END_IF;
   #IEC_Timer_1_Instance.TON(IN := #_w8 AND #Static05, PT := T#1000ms);
   IF #IEC_Timer_1_Instance.Q AND (#AdjustmentStatus = 2047) THEN #AdjustStep := #AdjustStep; END_IF;
   #_w9 := #IEC_Timer_1_Instance.Q AND (#AdjustmentStatus = 2045);
   #_w10 := #_w9 AND NOT #Static06;   // rising edge
   #Static06 := #_w9;
   IF #_w10 THEN
       #CurrentPoint_0 := #CurrentPoint_0 + 1;
       #AdjustStep := 4;
   END_IF;
   IF #IEC_Timer_1_Instance.Q AND (#AdjustmentStatus = 2046) THEN #AdjustStep := 6; END_IF;
   IF #IEC_Timer_1_Instance.Q AND (#AdjustmentStatus < 0) THEN #AdjustStep := 8; END_IF;
   #_w11 := #_w1 AND (#AdjustStep = 6);
   IF #_w11 THEN #Validate_REC := 1; END_IF;
   #WRREC_SpanAdjust.REQ := #_w11 AND NOT #WRREC_SpanAdjust.DONE;
   IF #_w11 THEN
       #WRREC_SpanAdjust(REQ := #WRREC_SpanAdjust.REQ,   // WRREC
                         ID := #ID,
                         INDEX := 16#4010,
                         LEN := 1,
                         RECORD := #Validate_REC,
                         DONE => #WRREC_SpanAdjust.DONE,
                         BUSY => #WRREC_SpanAdjust.BUSY,
                         ERROR => #WRREC_SpanAdjust.ERROR,
                         STATUS => #WRREC_SpanAdjust.STATUS);
   END_IF;
   #_w12 := #_w11 AND #WRREC_SpanAdjust.DONE AND NOT #Static07;   // rising edge of #WRREC_SpanAdjust.DONE
   #Static07 := #WRREC_SpanAdjust.DONE;
   IF #_w12 THEN #AdjustStep := 7; END_IF;
   IF #_w1 AND (#AdjustStep = 7) AND (#AdjustmentStatus = 0) THEN
       #CurrentPoint_0 := 0;
       #CurrentWeight_0 := 0.0;
       #Done := TRUE;
       #Error := FALSE;
       #Cancelled := FALSE;
       #Start := FALSE;
       #Static05 := FALSE;
       #Activate := FALSE;
       #AdjustStep := 0;
   END_IF;
   IF #_w1 AND (#AdjustStep = 8) THEN
       #CurrentPoint_0 := 0;
       #CurrentWeight_0 := 0.0;
       #Error := TRUE;
       #ConfirmWeight := FALSE;
       #Done := FALSE;
       #Cancelled := FALSE;
       #Start := FALSE;
       #Static05 := FALSE;
       #Activate := FALSE;
       #AdjustStep := 0;
   END_IF;
   #_w13 := #_w1 AND (#AdjustStep >= 4);
   #RDREC_Status.REQ := #_w13 AND NOT #RDREC_Status.VALID;
   IF #_w13 THEN
       #RDREC_Status(REQ := #RDREC_Status.REQ,   // RDREC
                     ID := #ID,
                     INDEX := 16#4007,
                     MLEN := 2,
                     RECORD := #AdjustmentStatus,
                     VALID => #RDREC_Status.VALID,
                     BUSY => #RDREC_Status.BUSY,
                     ERROR => #RDREC_Status.ERROR,
                     STATUS => #RDREC_Status.STATUS);
   END_IF;
END_REGION

REGION Network 3: Adjsutment Status
   // LoadWeight - Inform user to load the next adjustment weight according to CurrentWeight value
   // Process - Status bit to inform that the weight transmitter is performing adjustment process
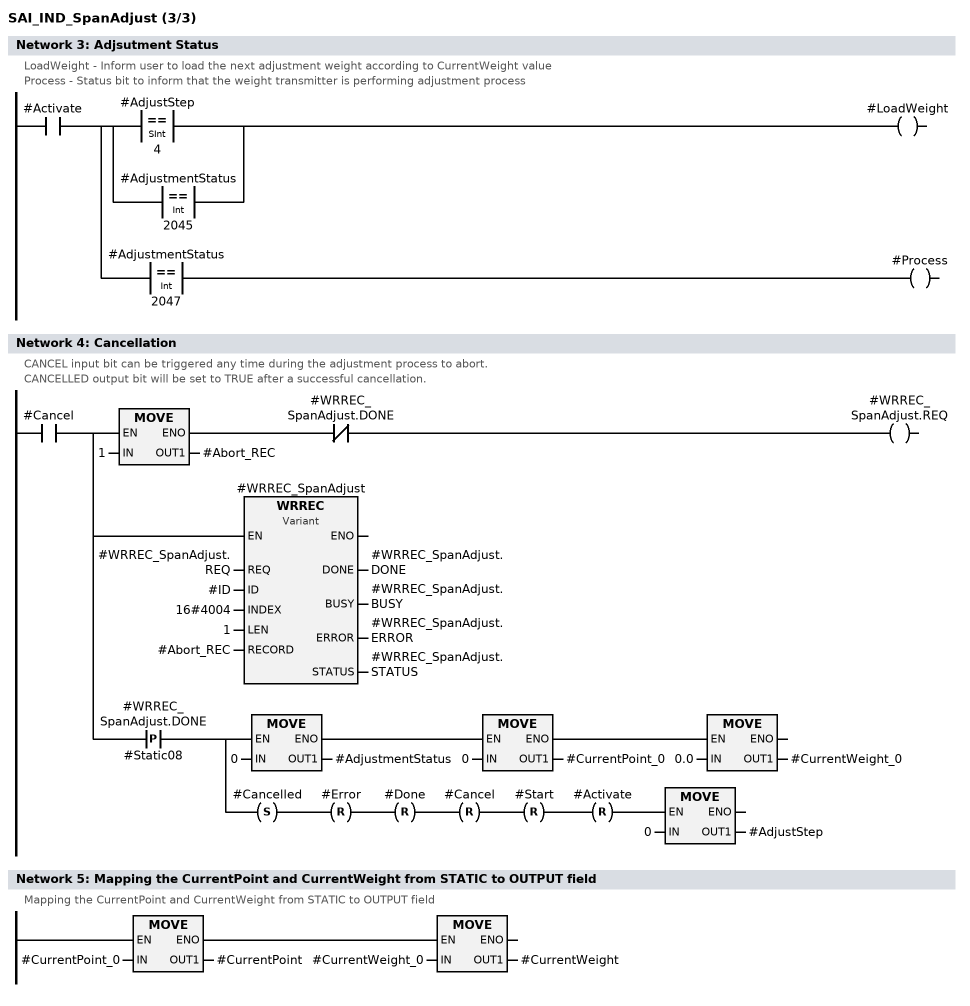
   RUNG wire#powerrail
      Contact( #Activate )
      wire#w1
      { S7_Templates := "SrcType := SInt" } EQ_Contact(in1 := #AdjustStep, in2 := 4)
      wire#w2
      Coil( #LoadWeight )
   END_RUNG
   RUNG wire#w1
      { S7_Templates := "SrcType := Int" } EQ_Contact(in1 := #AdjustmentStatus, in2 := 2045)
   END_RUNG wire#w2
   RUNG wire#w1
      { S7_Templates := "SrcType := Int" } EQ_Contact(in1 := #AdjustmentStatus, in2 := 2047)
      Coil( #Process )
   END_RUNG
   // the same network as SCL:
   #LoadWeight := #Activate AND ((#AdjustStep = 4) OR (#AdjustmentStatus = 2045));
   #Process := #Activate AND (#AdjustmentStatus = 2047);
END_REGION

REGION Network 4: Cancellation
   // CANCEL input bit can be triggered any time during the adjustment process to abort. 
   // CANCELLED output bit will be set to TRUE after a successful cancellation.
   RUNG wire#powerrail
      Contact( #Cancel )
      wire#w1
      Move(in := 1, out1 => #Abort_REC)
      I_Contact( #WRREC_SpanAdjust.DONE )
      Coil( #WRREC_SpanAdjust.REQ )
   END_RUNG
   RUNG wire#w1
      { S7_Templates := "[ptr_type := Variant, id_type := HW_IO, index_type := DInt, len_type := UInt]" } #WRREC_SpanAdjust.WRREC(REQ := #WRREC_SpanAdjust.REQ, ID := #ID, INDEX := 16#4004, LEN := 1, RECORD := #Abort_REC, DONE => #WRREC_SpanAdjust.DONE, BUSY => #WRREC_SpanAdjust.BUSY, ERROR => #WRREC_SpanAdjust.ERROR, STATUS => #WRREC_SpanAdjust.STATUS)
   END_RUNG
   RUNG wire#w1
      P_Contact(operand := #WRREC_SpanAdjust.DONE, bit := #Static08)
      wire#w2
      Move(in := 0, out1 => #AdjustmentStatus)
      Move(in := 0, out1 => #CurrentPoint_0)
      Move(in := 0.0, out1 => #CurrentWeight_0)
   END_RUNG
   RUNG wire#w2
      S_Coil( #Cancelled )
      R_Coil( #Error )
      R_Coil( #Done )
      R_Coil( #Cancel )
      R_Coil( #Start )
      R_Coil( #Activate )
      Move(in := 0, out1 => #AdjustStep)
   END_RUNG
   // the same network as SCL:
   IF #Cancel THEN #Abort_REC := 1; END_IF;
   #WRREC_SpanAdjust.REQ := #Cancel AND NOT #WRREC_SpanAdjust.DONE;
   IF #Cancel THEN
       #WRREC_SpanAdjust(REQ := #WRREC_SpanAdjust.REQ,   // WRREC
                         ID := #ID,
                         INDEX := 16#4004,
                         LEN := 1,
                         RECORD := #Abort_REC,
                         DONE => #WRREC_SpanAdjust.DONE,
                         BUSY => #WRREC_SpanAdjust.BUSY,
                         ERROR => #WRREC_SpanAdjust.ERROR,
                         STATUS => #WRREC_SpanAdjust.STATUS);
   END_IF;
   #_w1 := #Cancel AND #WRREC_SpanAdjust.DONE AND NOT #Static08;   // rising edge of #WRREC_SpanAdjust.DONE
   #Static08 := #WRREC_SpanAdjust.DONE;
   IF #_w1 THEN
       #AdjustmentStatus := 0;
       #CurrentPoint_0 := 0;
       #CurrentWeight_0 := 0.0;
       #Cancelled := TRUE;
       #Error := FALSE;
       #Done := FALSE;
       #Cancel := FALSE;
       #Start := FALSE;
       #Activate := FALSE;
       #AdjustStep := 0;
   END_IF;
END_REGION

REGION Network 5: Mapping the CurrentPoint and CurrentWeight from STATIC to OUTPUT field
   // Mapping the CurrentPoint and CurrentWeight from STATIC to OUTPUT field
   RUNG wire#powerrail
      Move(in := #CurrentPoint_0, out1 => #CurrentPoint)
      Move(in := #CurrentWeight_0, out1 => #CurrentWeight)
   END_RUNG
   // the same network as SCL:
   #CurrentPoint := #CurrentPoint_0;
   #CurrentWeight := #CurrentWeight_0;
END_REGION
END_FUNCTION_BLOCK

FUNCTION_BLOCK "SAI_IND_CalFree"   // FB53, LAD
TITLE = CalFree Adjustment
{ S7_Optimized_Access := 'FALSE' }
VERSION : 0.1
// CalFree is a method of analog scale adjustment without using test weights. It takes the factory calibrated load cell Rated Output (mV/ Vexc.) and user defined scale capacity to build a linear loading curve.
// This method is usually applied to huge capacity scales in which calibration with test weights or other material is not feasible at all.
// stored: AutoNumber true, IsIECCheckEnabled false, SetENOAutomatically false, UDAEnableTagReadback false
   VAR_INPUT
      ID : HW_IO;   // The Profinet Device Hardware Identifier under device properties
   END_VAR
   VAR_OUTPUT
      Process : Bool;   // Adjustment is in process
      Done : Bool;   // Adjustment completed successfully
      Error : Bool;
   END_VAR
   VAR_IN_OUT
      RatedCapacity : Real;   // Scale Capacity
      Unit : SInt := 1;   // Decimal 0 - gram; 1 - KG; 2 - Lbs
      RatedOutput : Real;   // The averaged load cells' Rated Output in mV/V
      Start : Bool;   // Switch ON to start adjustment
   END_VAR
   VAR DB_SPECIFIC
      Activate : Bool;
      Status_RECORD : Int;
      CalFree_RECORD : Int;
      AdjustStep : SInt;
      Check01 : Bool;
      Check02 : Bool;
   END_VAR
   VAR
      WRREC_CalFree { S7_SetPoint := 'True'} : WRREC;
   END_VAR
   VAR DB_SPECIFIC
      Static01 : Bool;
   END_VAR
   VAR
      RDREC_Status { S7_SetPoint := 'True'} : RDREC;
   END_VAR
   VAR_TEMP   // added for the SCL form of the ladder/FBD networks
      _w1 : Bool;
      _w2 : Bool;
      _w3 : Bool;
      _w4 : Bool;
      _w5 : Bool;
      _w6 : Bool;
      _w7 : Bool;
      _w8 : Bool;
      _w9 : Bool;
      _w10 : Bool;
      _w11 : Bool;
   END_VAR
BEGIN

REGION Network 1: Start routine
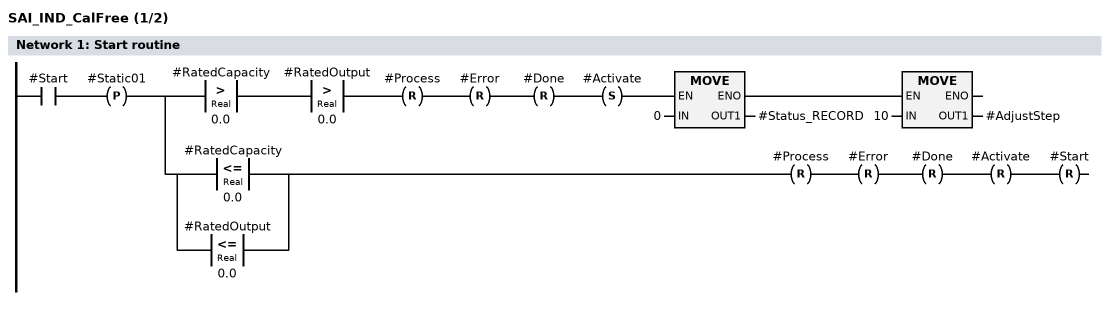
   RUNG wire#powerrail
      Contact( #Start )
      P_Trig( #Static01 )
      wire#w1
      { S7_Templates := "SrcType := Real" } GT_Contact(in1 := #RatedCapacity, in2 := 0.0)
      { S7_Templates := "SrcType := Real" } GT_Contact(in1 := #RatedOutput, in2 := 0.0)
      R_Coil( #Process )
      R_Coil( #Error )
      R_Coil( #Done )
      S_Coil( #Activate )
      Move(in := 0, out1 => #Status_RECORD)
      Move(in := 10, out1 => #AdjustStep)
   END_RUNG
   RUNG wire#w1
      { S7_Templates := "SrcType := Real" } LE_Contact(in1 := #RatedCapacity, in2 := 0.0)
      wire#w2
      R_Coil( #Process )
      R_Coil( #Error )
      R_Coil( #Done )
      R_Coil( #Activate )
      R_Coil( #Start )
   END_RUNG
   RUNG wire#w1
      { S7_Templates := "SrcType := Real" } LE_Contact(in1 := #RatedOutput, in2 := 0.0)
   END_RUNG wire#w2
   // the same network as SCL:
   #_w1 := #Start AND NOT #Static01;   // rising edge
   #Static01 := #Start;
   IF #_w1 AND (#RatedCapacity > 0.0) AND (#RatedOutput > 0.0) THEN
       #Process := FALSE;
       #Error := FALSE;
       #Done := FALSE;
       #Activate := TRUE;
       #Status_RECORD := 0;
       #AdjustStep := 10;
   END_IF;
   IF #_w1 AND ((#RatedCapacity <= 0.0) OR (#RatedOutput <= 0.0)) THEN
       #Process := FALSE;
       #Error := FALSE;
       #Done := FALSE;
       #Activate := FALSE;
       #Start := FALSE;
   END_IF;
END_REGION

REGION Network 2: Sequence
   // CalFree adjustment steps:
   // 
   // 1. Switch on Input bit Start
   // 
   // 2. Write in (a) Scale Capacity (Index 0x401A), (b) Scale unit (Index 0x401C, Decimal 0 - gram; Decimal 1 - KG; Decimal 2 - Pounds) and (c) Load Cells' averaged Rated Output (Index 0x401D, in mV/V)
   // 
   // 3. Start CalFree adjustment (Index 0x401A)
   // 
   // 4. Continuously read in adjustment status (Index 0x4007)
   // 
   // 5. Output bit Done will be turned ON after completion of the process
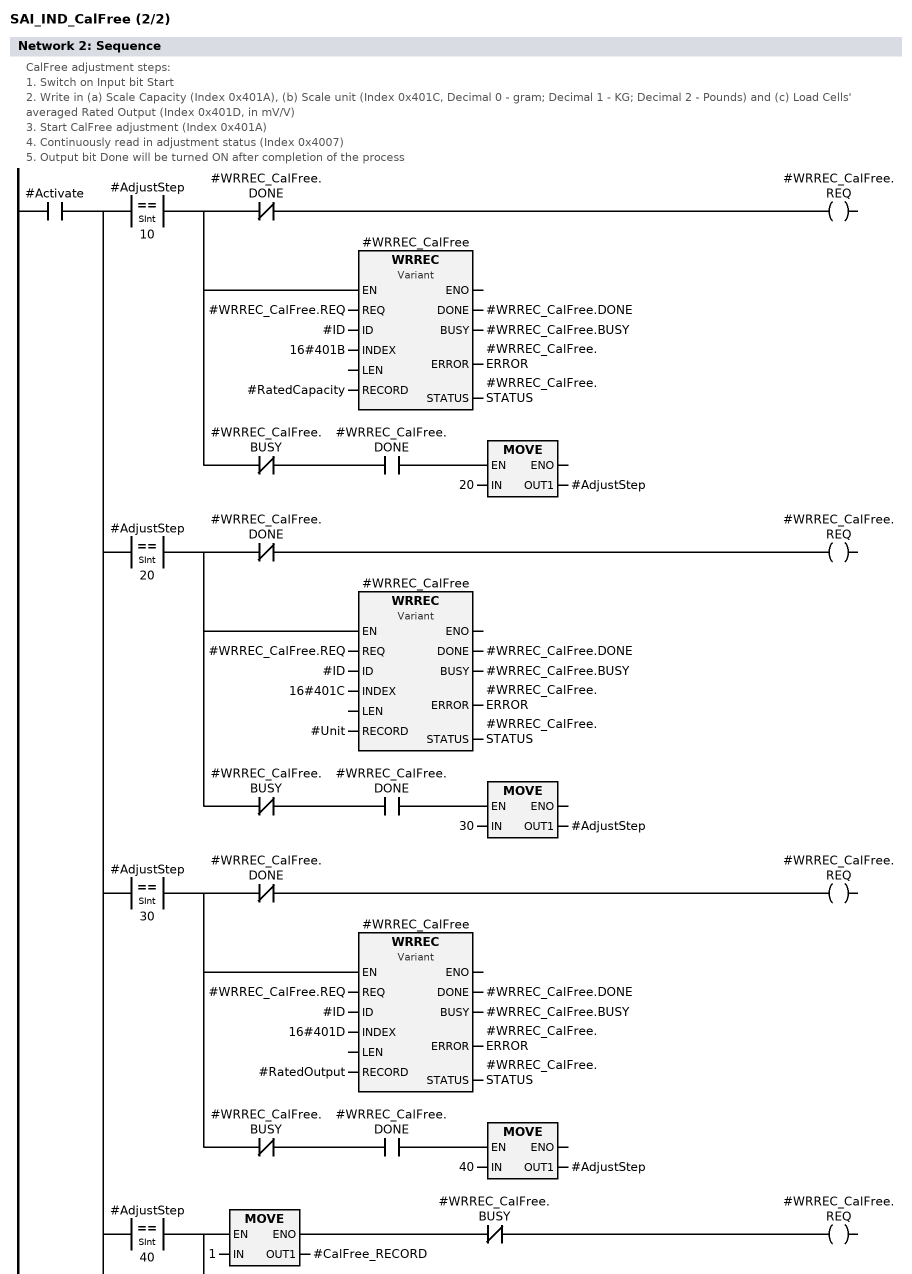
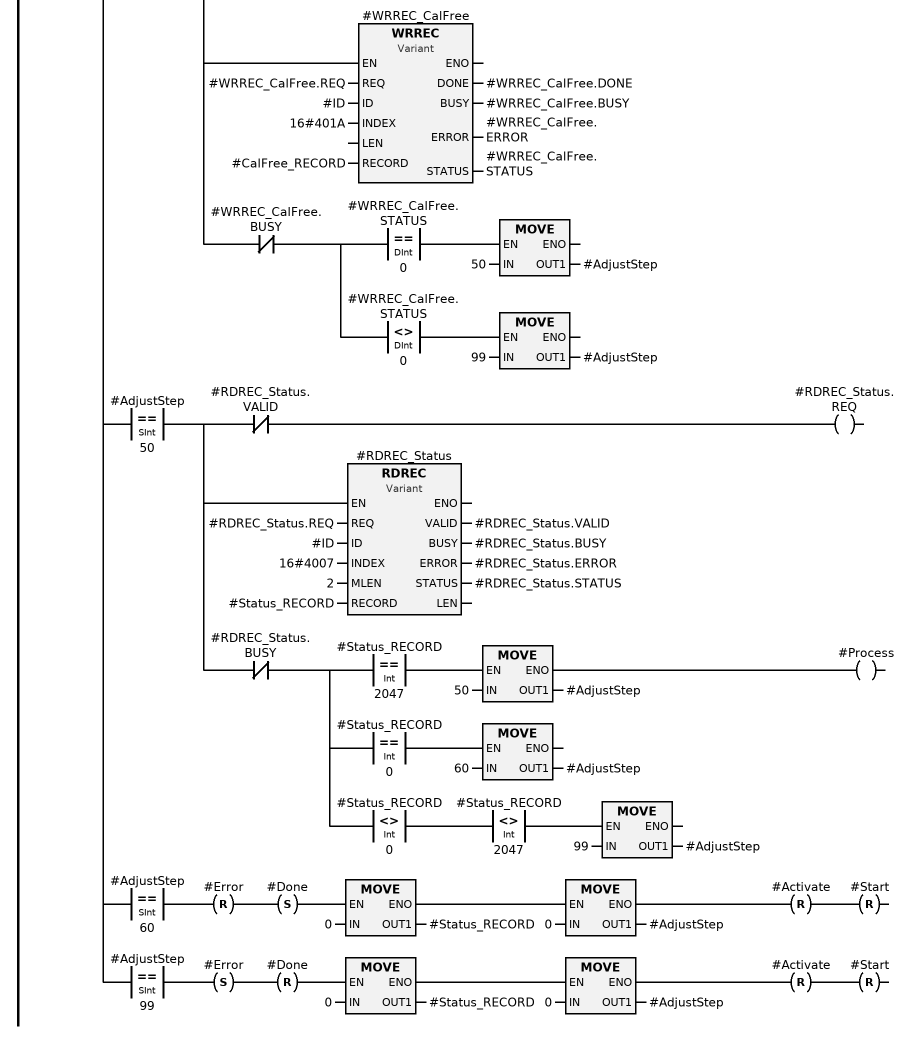
   RUNG wire#powerrail
      Contact( #Activate )
      wire#w1
      { S7_Templates := "SrcType := SInt" } EQ_Contact(in1 := #AdjustStep, in2 := 10)
      wire#w2
      I_Contact( #WRREC_CalFree.DONE )
      Coil( #WRREC_CalFree.REQ )
   END_RUNG
   RUNG wire#w2
      { S7_Templates := "[ptr_type := Variant, id_type := HW_IO, index_type := DInt, len_type := UInt]" } #WRREC_CalFree.WRREC(REQ := #WRREC_CalFree.REQ, ID := #ID, INDEX := 16#401B, LEN :=, RECORD := #RatedCapacity, DONE => #WRREC_CalFree.DONE, BUSY => #WRREC_CalFree.BUSY, ERROR => #WRREC_CalFree.ERROR, STATUS => #WRREC_CalFree.STATUS)
   END_RUNG
   RUNG wire#w2
      I_Contact( #WRREC_CalFree.BUSY )
      Contact( #WRREC_CalFree.DONE )
      Move(in := 20, out1 => #AdjustStep)
   END_RUNG
   RUNG wire#w1
      { S7_Templates := "SrcType := SInt" } EQ_Contact(in1 := #AdjustStep, in2 := 20)
      wire#w3
      I_Contact( #WRREC_CalFree.DONE )
      Coil( #WRREC_CalFree.REQ )
   END_RUNG
   RUNG wire#w3
      { S7_Templates := "[ptr_type := Variant, id_type := HW_IO, index_type := DInt, len_type := UInt]" } #WRREC_CalFree.WRREC(REQ := #WRREC_CalFree.REQ, ID := #ID, INDEX := 16#401C, LEN :=, RECORD := #Unit, DONE => #WRREC_CalFree.DONE, BUSY => #WRREC_CalFree.BUSY, ERROR => #WRREC_CalFree.ERROR, STATUS => #WRREC_CalFree.STATUS)
   END_RUNG
   RUNG wire#w3
      I_Contact( #WRREC_CalFree.BUSY )
      Contact( #WRREC_CalFree.DONE )
      Move(in := 30, out1 => #AdjustStep)
   END_RUNG
   RUNG wire#w1
      { S7_Templates := "SrcType := SInt" } EQ_Contact(in1 := #AdjustStep, in2 := 30)
      wire#w4
      I_Contact( #WRREC_CalFree.DONE )
      Coil( #WRREC_CalFree.REQ )
   END_RUNG
   RUNG wire#w4
      { S7_Templates := "[ptr_type := Variant, id_type := HW_IO, index_type := DInt, len_type := UInt]" } #WRREC_CalFree.WRREC(REQ := #WRREC_CalFree.REQ, ID := #ID, INDEX := 16#401D, LEN :=, RECORD := #RatedOutput, DONE => #WRREC_CalFree.DONE, BUSY => #WRREC_CalFree.BUSY, ERROR => #WRREC_CalFree.ERROR, STATUS => #WRREC_CalFree.STATUS)
   END_RUNG
   RUNG wire#w4
      I_Contact( #WRREC_CalFree.BUSY )
      Contact( #WRREC_CalFree.DONE )
      Move(in := 40, out1 => #AdjustStep)
   END_RUNG
   RUNG wire#w1
      { S7_Templates := "SrcType := SInt" } EQ_Contact(in1 := #AdjustStep, in2 := 40)
      wire#w5
      Move(in := 1, out1 => #CalFree_RECORD)
      I_Contact( #WRREC_CalFree.BUSY )
      Coil( #WRREC_CalFree.REQ )
   END_RUNG
   RUNG wire#w5
      { S7_Templates := "[ptr_type := Variant, id_type := HW_IO, index_type := DInt, len_type := UInt]" } #WRREC_CalFree.WRREC(REQ := #WRREC_CalFree.REQ, ID := #ID, INDEX := 16#401A, LEN :=, RECORD := #CalFree_RECORD, DONE => #WRREC_CalFree.DONE, BUSY => #WRREC_CalFree.BUSY, ERROR => #WRREC_CalFree.ERROR, STATUS => #WRREC_CalFree.STATUS)
   END_RUNG
   RUNG wire#w5
      I_Contact( #WRREC_CalFree.BUSY )
      wire#w6
      { S7_Templates := "SrcType := DInt" } EQ_Contact(in1 := #WRREC_CalFree.STATUS, in2 := 0)
      Move(in := 50, out1 => #AdjustStep)
   END_RUNG
   RUNG wire#w6
      { S7_Templates := "SrcType := DInt" } NE_Contact(in1 := #WRREC_CalFree.STATUS, in2 := 0)
      Move(in := 99, out1 => #AdjustStep)
   END_RUNG
   RUNG wire#w1
      { S7_Templates := "SrcType := SInt" } EQ_Contact(in1 := #AdjustStep, in2 := 50)
      wire#w7
      I_Contact( #RDREC_Status.VALID )
      Coil( #RDREC_Status.REQ )
   END_RUNG
   RUNG wire#w7
      { S7_Templates := "[ptr_type := Variant, id_type := HW_IO, index_type := DInt, len_type := UInt]" } #RDREC_Status.RDREC(REQ := #RDREC_Status.REQ, ID := #ID, INDEX := 16#4007, MLEN := 2, RECORD := #Status_RECORD, VALID => #RDREC_Status.VALID, BUSY => #RDREC_Status.BUSY, ERROR => #RDREC_Status.ERROR, STATUS => #RDREC_Status.STATUS, LEN =>)
   END_RUNG
   RUNG wire#w7
      I_Contact( #RDREC_Status.BUSY )
      wire#w8
      { S7_Templates := "SrcType := Int" } EQ_Contact(in1 := #Status_RECORD, in2 := 2047)
      Move(in := 50, out1 => #AdjustStep)
      Coil( #Process )
   END_RUNG
   RUNG wire#w8
      { S7_Templates := "SrcType := Int" } EQ_Contact(in1 := #Status_RECORD, in2 := 0)
      Move(in := 60, out1 => #AdjustStep)
   END_RUNG
   RUNG wire#w8
      { S7_Templates := "SrcType := Int" } NE_Contact(in1 := #Status_RECORD, in2 := 0)
      { S7_Templates := "SrcType := Int" } NE_Contact(in1 := #Status_RECORD, in2 := 2047)
      Move(in := 99, out1 => #AdjustStep)
   END_RUNG
   RUNG wire#w1
      { S7_Templates := "SrcType := SInt" } EQ_Contact(in1 := #AdjustStep, in2 := 60)
      R_Coil( #Error )
      S_Coil( #Done )
      Move(in := 0, out1 => #Status_RECORD)
      Move(in := 0, out1 => #AdjustStep)
      R_Coil( #Activate )
      R_Coil( #Start )
   END_RUNG
   RUNG wire#w1
      { S7_Templates := "SrcType := SInt" } EQ_Contact(in1 := #AdjustStep, in2 := 99)
      S_Coil( #Error )
      R_Coil( #Done )
      Move(in := 0, out1 => #Status_RECORD)
      Move(in := 0, out1 => #AdjustStep)
      R_Coil( #Activate )
      R_Coil( #Start )
   END_RUNG
   // the same network as SCL:
   #_w1 := #Activate AND (#AdjustStep = 10);
   #WRREC_CalFree.REQ := #_w1 AND NOT #WRREC_CalFree.DONE;
   IF #_w1 THEN
       #WRREC_CalFree(REQ := #WRREC_CalFree.REQ,   // WRREC
                      ID := #ID,
                      INDEX := 16#401B,
                      RECORD := #RatedCapacity,
                      DONE => #WRREC_CalFree.DONE,
                      BUSY => #WRREC_CalFree.BUSY,
                      ERROR => #WRREC_CalFree.ERROR,
                      STATUS => #WRREC_CalFree.STATUS);
   END_IF;
   IF #_w1 AND NOT #WRREC_CalFree.BUSY AND #WRREC_CalFree.DONE THEN #AdjustStep := 20; END_IF;
   #_w2 := #Activate AND (#AdjustStep = 20);
   #WRREC_CalFree.REQ := #_w2 AND NOT #WRREC_CalFree.DONE;
   IF #_w2 THEN
       #WRREC_CalFree(REQ := #WRREC_CalFree.REQ,   // WRREC
                      ID := #ID,
                      INDEX := 16#401C,
                      RECORD := #Unit,
                      DONE => #WRREC_CalFree.DONE,
                      BUSY => #WRREC_CalFree.BUSY,
                      ERROR => #WRREC_CalFree.ERROR,
                      STATUS => #WRREC_CalFree.STATUS);
   END_IF;
   IF #_w2 AND NOT #WRREC_CalFree.BUSY AND #WRREC_CalFree.DONE THEN #AdjustStep := 30; END_IF;
   #_w3 := #Activate AND (#AdjustStep = 30);
   #WRREC_CalFree.REQ := #_w3 AND NOT #WRREC_CalFree.DONE;
   IF #_w3 THEN
       #WRREC_CalFree(REQ := #WRREC_CalFree.REQ,   // WRREC
                      ID := #ID,
                      INDEX := 16#401D,
                      RECORD := #RatedOutput,
                      DONE => #WRREC_CalFree.DONE,
                      BUSY => #WRREC_CalFree.BUSY,
                      ERROR => #WRREC_CalFree.ERROR,
                      STATUS => #WRREC_CalFree.STATUS);
   END_IF;
   IF #_w3 AND NOT #WRREC_CalFree.BUSY AND #WRREC_CalFree.DONE THEN #AdjustStep := 40; END_IF;
   #_w4 := #Activate AND (#AdjustStep = 40);
   IF #_w4 THEN #CalFree_RECORD := 1; END_IF;
   #WRREC_CalFree.REQ := #_w4 AND NOT #WRREC_CalFree.BUSY;
   IF #_w4 THEN
       #WRREC_CalFree(REQ := #WRREC_CalFree.REQ,   // WRREC
                      ID := #ID,
                      INDEX := 16#401A,
                      RECORD := #CalFree_RECORD,
                      DONE => #WRREC_CalFree.DONE,
                      BUSY => #WRREC_CalFree.BUSY,
                      ERROR => #WRREC_CalFree.ERROR,
                      STATUS => #WRREC_CalFree.STATUS);
   END_IF;
   #_w5 := #_w4 AND NOT #WRREC_CalFree.BUSY;
   IF #_w5 AND (#WRREC_CalFree.STATUS = 0) THEN #AdjustStep := 50; END_IF;
   IF #_w5 AND (#WRREC_CalFree.STATUS <> 0) THEN #AdjustStep := 99; END_IF;
   #_w6 := #Activate AND (#AdjustStep = 50);
   #RDREC_Status.REQ := #_w6 AND NOT #RDREC_Status.VALID;
   IF #_w6 THEN
       #RDREC_Status(REQ := #RDREC_Status.REQ,   // RDREC
                     ID := #ID,
                     INDEX := 16#4007,
                     MLEN := 2,
                     RECORD := #Status_RECORD,
                     VALID => #RDREC_Status.VALID,
                     BUSY => #RDREC_Status.BUSY,
                     ERROR => #RDREC_Status.ERROR,
                     STATUS => #RDREC_Status.STATUS);
   END_IF;
   #_w7 := #_w6 AND NOT #RDREC_Status.BUSY;
   #_w8 := #_w7 AND (#Status_RECORD = 2047);
   IF #_w8 THEN #AdjustStep := 50; END_IF;
   #Process := #_w8;
   IF #_w7 AND (#Status_RECORD = 0) THEN #AdjustStep := 60; END_IF;
   IF #_w7 AND (#Status_RECORD <> 0) AND (#Status_RECORD <> 2047) THEN #AdjustStep := 99; END_IF;
   IF #Activate AND (#AdjustStep = 60) THEN
       #Error := FALSE;
       #Done := TRUE;
       #Status_RECORD := 0;
   END_IF;
   #_w9 := #Activate AND (#AdjustStep = 60);
   IF #_w9 THEN #AdjustStep := 0; END_IF;
   #_w10 := #Activate;
   IF #_w9 THEN
       #Activate := FALSE;
       #Start := FALSE;
   END_IF;
   IF #_w10 AND (#AdjustStep = 99) THEN
       #Error := TRUE;
       #Done := FALSE;
       #Status_RECORD := 0;
   END_IF;
   #_w11 := #_w10 AND (#AdjustStep = 99);
   IF #_w11 THEN
       #AdjustStep := 0;
       #Activate := FALSE;
       #Start := FALSE;
   END_IF;
END_REGION
END_FUNCTION_BLOCK

FUNCTION_BLOCK "SAI_IND360Base_AlibiRead"   // FB4, LAD
{ S7_Optimized_Access := 'FALSE' }
VERSION : 0.1
// stored: AutoNumber true, IsIECCheckEnabled false, SetENOAutomatically false, UDAEnableTagReadback false
   VAR_INPUT
      ID : HW_IO;   // The Profinet Device Hardware Identifier under device properties
   END_VAR
   VAR_OUTPUT
      Done : Bool;   // Read done successfully
      Error : Bool;   // Error during reading process
      GrossWeight : Real;
      TareWeight : Real;
      NetWeight : Real;
      TareMode : SInt;   // 0,tare;1;preset tare
      Unit : SInt;   // Unit: 0-g; 1-kg, 2-lb
   END_VAR
   VAR_IN_OUT
      ePrint : Bool;   // Toggle this bit to execute an ePrint from terminal > PLC
      RecordNumber : DInt;   // record number which is to be read out from the weighing indicator
      Get_TransactionNum : Bool;   // Trigger this bit to get the previously read alibi record number.
      Set_TransactionNum : Bool;   // Trigger this bit to set the alibi record number which is to be read out
      Get_Alibi : Bool;   // Trigger this bit to read out the alibi transaction record specified by "RecordNum".
      Alibi_Array : Array[0..44] of Byte;
   END_VAR
   VAR
      RDREC01 { S7_SetPoint := 'True'} : RDREC;
      RDREC02 { S7_SetPoint := 'True'} : RDREC;
      WRREC01 { S7_SetPoint := 'True'} : WRREC;
      WRREC02 { S7_SetPoint := 'True'} : WRREC;
   END_VAR
   VAR DB_SPECIFIC
      UINT : SInt;
   END_VAR
BEGIN

REGION Network 1: Read transaction number
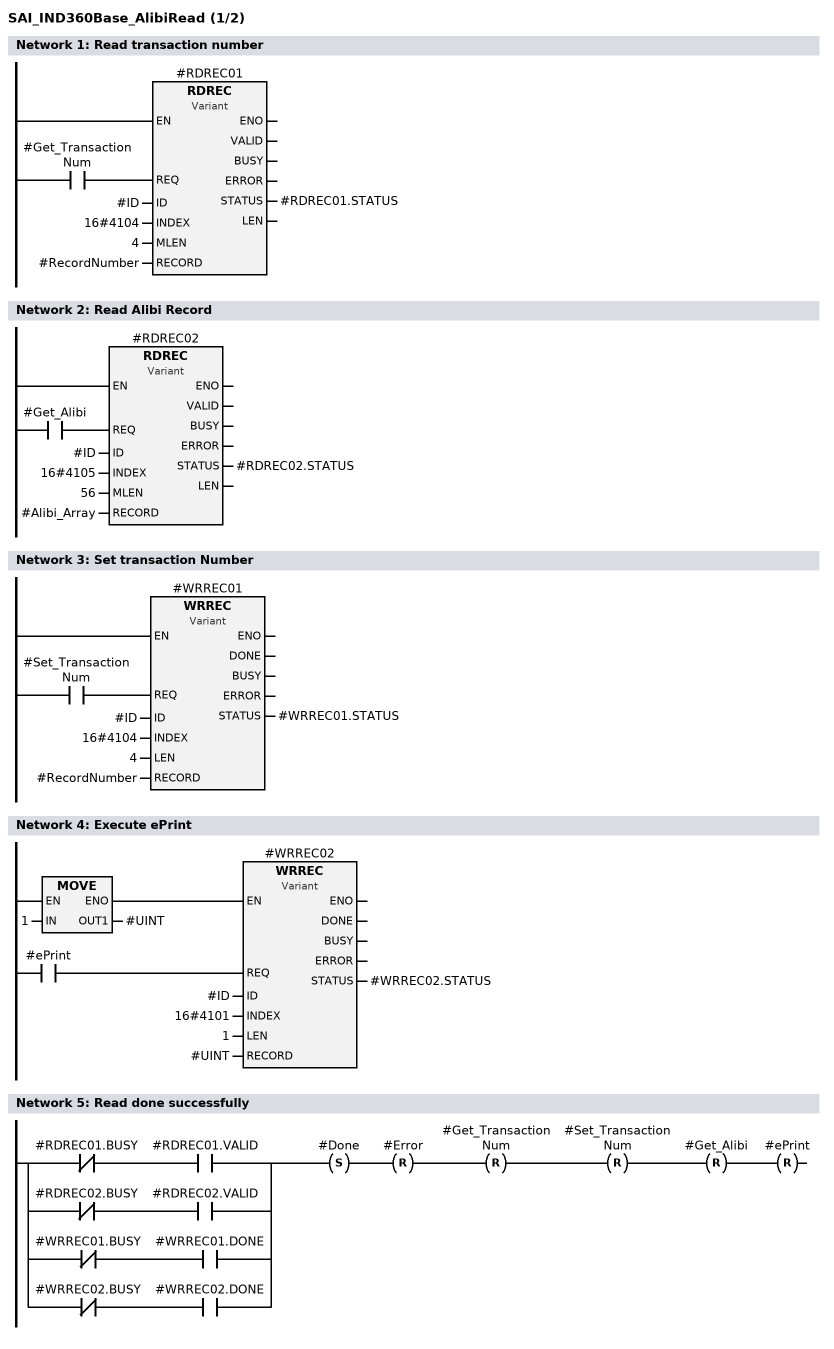
   RUNG wire#powerrail
      { S7_Templates := "[ptr_type := Variant, id_type := HW_IO, index_type := DInt, len_type := UInt]" } #RDREC01.RDREC(REQ := wire#w1, ID := #ID, INDEX := 16#4104, MLEN := 4, RECORD := #RecordNumber, VALID =>, BUSY =>, ERROR =>, STATUS => #RDREC01.STATUS, LEN =>)
   END_RUNG
   RUNG wire#powerrail
      Contact( #Get_TransactionNum )
   END_RUNG wire#w1
   // the same network as SCL:
   #RDREC01(REQ := #Get_TransactionNum,   // RDREC
            ID := #ID,
            INDEX := 16#4104,
            MLEN := 4,
            RECORD := #RecordNumber,
            STATUS => #RDREC01.STATUS);
END_REGION

REGION Network 2: Read Alibi Record
   RUNG wire#powerrail
      { S7_Templates := "[ptr_type := Variant, id_type := HW_IO, index_type := DInt, len_type := UInt]" } #RDREC02.RDREC(REQ := wire#w1, ID := #ID, INDEX := 16#4105, MLEN := 56, RECORD := #Alibi_Array, VALID =>, BUSY =>, ERROR =>, STATUS => #RDREC02.STATUS, LEN =>)
   END_RUNG
   RUNG wire#powerrail
      Contact( #Get_Alibi )
   END_RUNG wire#w1
   // the same network as SCL:
   #RDREC02(REQ := #Get_Alibi,   // RDREC
            ID := #ID,
            INDEX := 16#4105,
            MLEN := 56,
            RECORD := #Alibi_Array,
            STATUS => #RDREC02.STATUS);
END_REGION

REGION Network 3: Set transaction Number
   RUNG wire#powerrail
      { S7_Templates := "[ptr_type := Variant, id_type := HW_IO, index_type := DInt, len_type := UInt]" } #WRREC01.WRREC(REQ := wire#w1, ID := #ID, INDEX := 16#4104, LEN := 4, RECORD := #RecordNumber, DONE =>, BUSY =>, ERROR =>, STATUS => #WRREC01.STATUS)
   END_RUNG
   RUNG wire#powerrail
      Contact( #Set_TransactionNum )
   END_RUNG wire#w1
   // the same network as SCL:
   #WRREC01(REQ := #Set_TransactionNum,   // WRREC
            ID := #ID,
            INDEX := 16#4104,
            LEN := 4,
            RECORD := #RecordNumber,
            STATUS => #WRREC01.STATUS);
END_REGION

REGION Network 4: Execute ePrint
   RUNG wire#powerrail
      Move(in := 1, out1 => #UINT)
      { S7_Templates := "[ptr_type := Variant, id_type := HW_IO, index_type := DInt, len_type := UInt]" } #WRREC02.WRREC(REQ := wire#w1, ID := #ID, INDEX := 16#4101, LEN := 1, RECORD := #UINT, DONE =>, BUSY =>, ERROR =>, STATUS => #WRREC02.STATUS)
   END_RUNG
   RUNG wire#powerrail
      Contact( #ePrint )
   END_RUNG wire#w1
   // the same network as SCL:
   #UINT := 1;
   #WRREC02(REQ := #ePrint, ID := #ID, INDEX := 16#4101, LEN := 1, RECORD := #UINT, STATUS => #WRREC02.STATUS);   // WRREC
END_REGION

REGION Network 5: Read done successfully
   RUNG wire#powerrail
      I_Contact( #RDREC01.BUSY )
      Contact( #RDREC01.VALID )
      wire#w1
      S_Coil( #Done )
      R_Coil( #Error )
      R_Coil( #Get_TransactionNum )
      R_Coil( #Set_TransactionNum )
      R_Coil( #Get_Alibi )
      R_Coil( #ePrint )
   END_RUNG
   RUNG wire#powerrail
      I_Contact( #RDREC02.BUSY )
      Contact( #RDREC02.VALID )
   END_RUNG wire#w1
   RUNG wire#powerrail
      I_Contact( #WRREC01.BUSY )
      Contact( #WRREC01.DONE )
   END_RUNG wire#w1
   RUNG wire#powerrail
      I_Contact( #WRREC02.BUSY )
      Contact( #WRREC02.DONE )
   END_RUNG wire#w1
   // the same network as SCL:
   IF (NOT #RDREC01.BUSY AND #RDREC01.VALID) OR (NOT #RDREC02.BUSY AND #RDREC02.VALID) OR (NOT #WRREC01.BUSY AND #WRREC01.DONE) OR (NOT #WRREC02.BUSY AND #WRREC02.DONE) THEN
       #Done := TRUE;
       #Error := FALSE;
       #Get_TransactionNum := FALSE;
       #Set_TransactionNum := FALSE;
       #Get_Alibi := FALSE;
       #ePrint := FALSE;
   END_IF;
END_REGION

REGION Network 6: Read failed
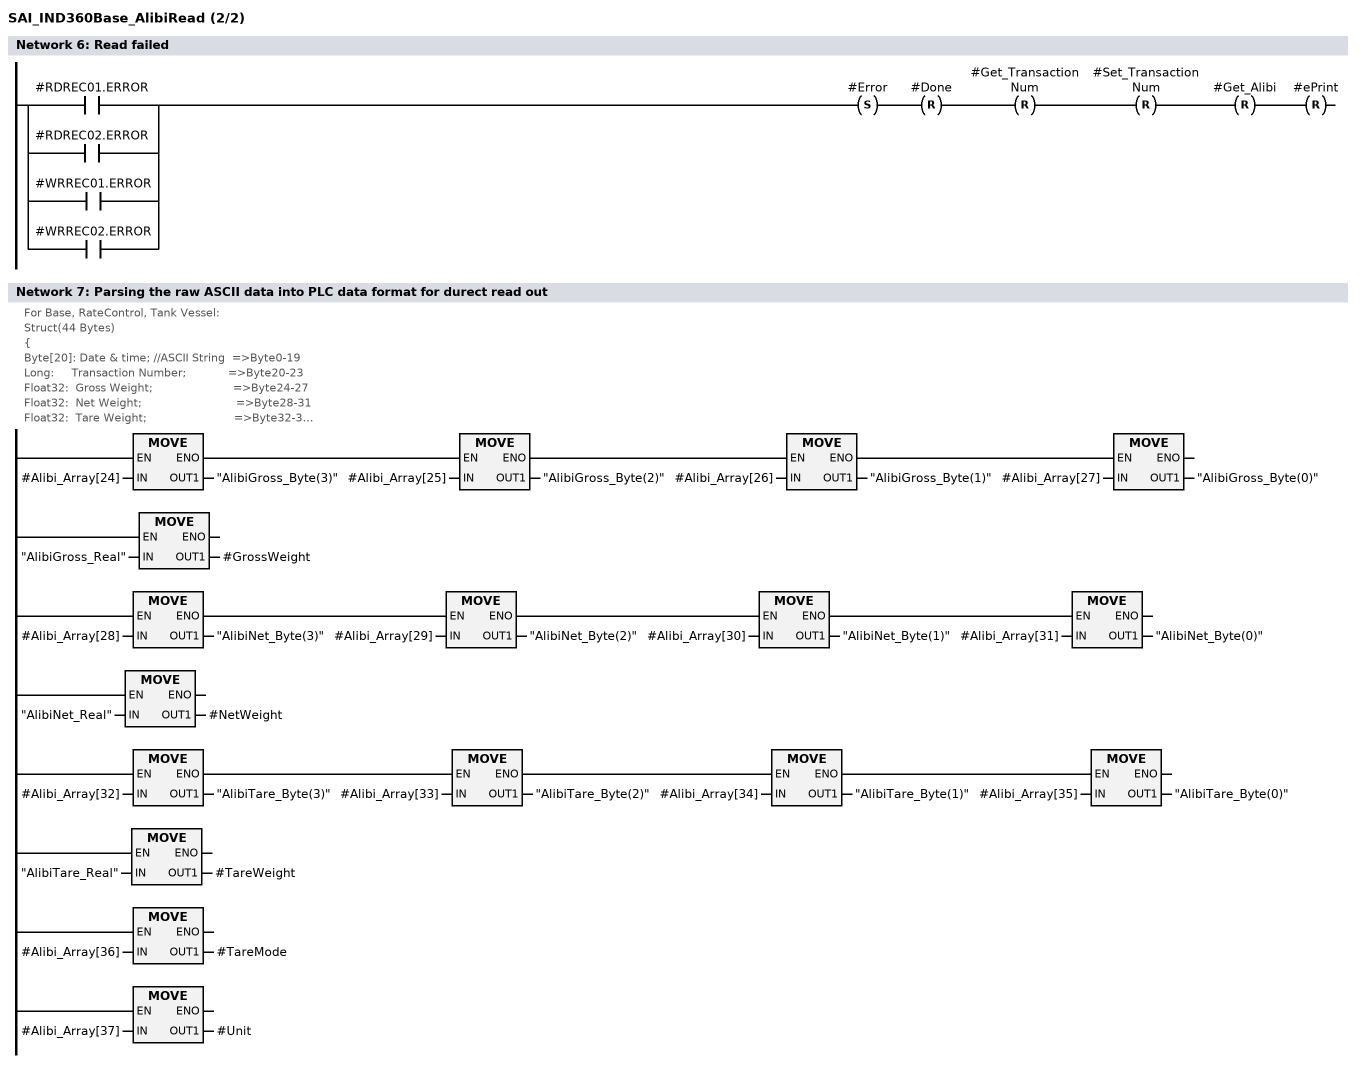
   RUNG wire#powerrail
      Contact( #RDREC01.ERROR )
      wire#w1
      S_Coil( #Error )
      R_Coil( #Done )
      R_Coil( #Get_TransactionNum )
      R_Coil( #Set_TransactionNum )
      R_Coil( #Get_Alibi )
      R_Coil( #ePrint )
   END_RUNG
   RUNG wire#powerrail
      Contact( #RDREC02.ERROR )
   END_RUNG wire#w1
   RUNG wire#powerrail
      Contact( #WRREC01.ERROR )
   END_RUNG wire#w1
   RUNG wire#powerrail
      Contact( #WRREC02.ERROR )
   END_RUNG wire#w1
   // the same network as SCL:
   IF #RDREC01.ERROR OR #RDREC02.ERROR OR #WRREC01.ERROR OR #WRREC02.ERROR THEN
       #Error := TRUE;
       #Done := FALSE;
       #Get_TransactionNum := FALSE;
       #Set_TransactionNum := FALSE;
       #Get_Alibi := FALSE;
       #ePrint := FALSE;
   END_IF;
END_REGION

REGION Network 7: Parsing the raw ASCII data into PLC data format for durect read out
   // For Base, RateControl, Tank Vessel:
   // Struct(44 Bytes)
   // {
   // Byte[20]: Date & time; //ASCII String  =>Byte0-19
   // Long:     Transaction Number;            =>Byte20-23
   // Float32:  Gross Weight;                       =>Byte24-27
   // Float32:  Net Weight;                           =>Byte28-31
   // Float32:  Tare Weight;                         =>Byte32-35
   // Byte:     Tare Mode;                              =>Byte36
   // Byte:     Unit;                                          =>Byte37
   // Byte[6]:  Not Used;                              =>Byte38-43
   // }
   RUNG wire#powerrail
      Move(in := #Alibi_Array[24], out1 => "AlibiGross_Byte(3)")
      Move(in := #Alibi_Array[25], out1 => "AlibiGross_Byte(2)")
      Move(in := #Alibi_Array[26], out1 => "AlibiGross_Byte(1)")
      Move(in := #Alibi_Array[27], out1 => "AlibiGross_Byte(0)")
   END_RUNG
   RUNG wire#powerrail
      Move(in := "AlibiGross_Real", out1 => #GrossWeight)
   END_RUNG
   RUNG wire#powerrail
      Move(in := #Alibi_Array[28], out1 => "AlibiNet_Byte(3)")
      Move(in := #Alibi_Array[29], out1 => "AlibiNet_Byte(2)")
      Move(in := #Alibi_Array[30], out1 => "AlibiNet_Byte(1)")
      Move(in := #Alibi_Array[31], out1 => "AlibiNet_Byte(0)")
   END_RUNG
   RUNG wire#powerrail
      Move(in := "AlibiNet_Real", out1 => #NetWeight)
   END_RUNG
   RUNG wire#powerrail
      Move(in := #Alibi_Array[32], out1 => "AlibiTare_Byte(3)")
      Move(in := #Alibi_Array[33], out1 => "AlibiTare_Byte(2)")
      Move(in := #Alibi_Array[34], out1 => "AlibiTare_Byte(1)")
      Move(in := #Alibi_Array[35], out1 => "AlibiTare_Byte(0)")
   END_RUNG
   RUNG wire#powerrail
      Move(in := "AlibiTare_Real", out1 => #TareWeight)
   END_RUNG
   RUNG wire#powerrail
      Move(in := #Alibi_Array[36], out1 => #TareMode)
   END_RUNG
   RUNG wire#powerrail
      Move(in := #Alibi_Array[37], out1 => #Unit)
   END_RUNG
   // the same network as SCL:
   "AlibiGross_Byte(3)" := #Alibi_Array[24];
   "AlibiGross_Byte(2)" := #Alibi_Array[25];
   "AlibiGross_Byte(1)" := #Alibi_Array[26];
   "AlibiGross_Byte(0)" := #Alibi_Array[27];
   #GrossWeight := "AlibiGross_Real";
   "AlibiNet_Byte(3)" := #Alibi_Array[28];
   "AlibiNet_Byte(2)" := #Alibi_Array[29];
   "AlibiNet_Byte(1)" := #Alibi_Array[30];
   "AlibiNet_Byte(0)" := #Alibi_Array[31];
   #NetWeight := "AlibiNet_Real";
   "AlibiTare_Byte(3)" := #Alibi_Array[32];
   "AlibiTare_Byte(2)" := #Alibi_Array[33];
   "AlibiTare_Byte(1)" := #Alibi_Array[34];
   "AlibiTare_Byte(0)" := #Alibi_Array[35];
   #TareWeight := "AlibiTare_Real";
   #TareMode := #Alibi_Array[36];
   #Unit := #Alibi_Array[37];
END_REGION
END_FUNCTION_BLOCK

FUNCTION "Profile Station FC" : Void   // FC32, SCL
{ S7_Optimized_Access := 'TRUE' }
VERSION : 0.1
// stored: AutoNumber true, IsIECCheckEnabled false, SetENOAutomatically false, UDAEnableTagReadback false
   VAR_INPUT
      MaxLength : Real;
      ConveyorSpeed_mm_s : Real;
   END_VAR
BEGIN
   "R_TRIG_DB_26"(CLK:="Control_DB"."Profiling Station".Start);

    "R_TRIG_DB_27"(CLK:=NOT "Profile Station - Cross 1" AND NOT "Profile Station - Cross 2",Q => "SensorUp");

    "IEC_Timer_0_DB_3".TON(IN:="Profile Station - Cross 1" AND "Profile Station - Cross 2",
                           PT:=T#2s,Q=>"SensorDown");


   CASE "State_PS" OF

           //-------------------------------------------------
           // 0 - IDLE
           //-------------------------------------------------
       0:
           "Control_DB"."Profiling Station".Error_ID := 0;
           "Control_DB"."Profiling Station".Ready := TRUE;
           "Control_DB"."Profiling Station".Running := FALSE;
           IF "R_TRIG_DB_26".Q THEN
               "Control_DB"."Profiling Station".Ready := FALSE;
               "Control_DB"."Profiling Station".Done := FALSE;
               "Control_DB"."Profiling Station".Valid := FALSE;
               "Control_DB"."Profiling Station".OverWidth := FALSE;
               "Control_DB"."Profiling Station".OverHeight := FALSE;
               "Control_DB"."Profiling Station".OverLength := FALSE;
               "Control_DB"."Profiling Station".Error_ID := 0;
               "Control_DB"."Profiling Station".Running := TRUE;
               "State_PS" := 10;
           END_IF;

       10:
           IF "SensorUp" THEN
               "State_PS" := 20;
           END_IF;

       20:
           "LengthTimer".TON(IN := TRUE,
                             PT := T#60S);

           IF NOT "Profile Station - Left" OR NOT "Profile Station - Right" THEN
               "Control_DB"."Profiling Station".OverWidth := TRUE;
           END_IF;

           IF NOT "Profile Station - High" THEN
               "Control_DB"."Profiling Station".OverHeight := TRUE;
           END_IF;

           IF "SensorDown" THEN
               "MeasuredTime_s" := DINT_TO_REAL(TIME_TO_DINT("LengthTimer".ET)) / 1000.0;
               "CalculatedLength" := "MeasuredTime_s" * #ConveyorSpeed_mm_s;

               // IF "CalculatedLength" > #MaxLength THEN
               //     "Control_DB"."Profiling Station".OverLength := TRUE;
               // END_IF;

               // Resultado final
               IF "Control_DB"."Profiling Station".OverWidth OR "Control_DB"."Profiling Station".OverHeight OR "Control_DB"."Profiling Station".OverLength THEN
                   "Control_DB"."Profiling Station".Valid := FALSE;
                   "Control_DB"."Profiling Station".Error_ID.%X0 := 1;
               ELSE
                   "Control_DB"."Profiling Station".Valid := TRUE;
                   "Control_DB"."Profiling Station".Error_ID := 0;
               END_IF;

               "LengthTimer".TON(IN := FALSE,
                                 PT := T#0S);
               "State_PS" := 100;
           END_IF;

       100:
           "Control_DB"."Profiling Station".Running := FALSE;
               "Control_DB"."Profiling Station".Done := TRUE;
               "State_PS" := 0;


       END_CASE;

       "IEC_Timer_0_DB_12".TON(IN:="Control_DB"."Profiling Station".Running,
                               PT:=t#30s);

       IF "IEC_Timer_0_DB_12".Q THEN
           "Control_DB"."Profiling Station".Valid := FALSE;
           "Control_DB"."Profiling Station".Error_ID := 1;
           "State_PS" := 100;
       END_IF;
END_FUNCTION

FUNCTION_BLOCK "Barcode_Station_FB"   // FB33, SCL
{ S7_Optimized_Access := 'TRUE' }
VERSION : 0.1
// stored: AutoNumber true, IsIECCheckEnabled false, IsRetainMemResEnabled false, MemoryReserve 100, SetENOAutomatically false, UDAEnableTagReadback false
   VAR_INPUT
      Start : Bool;
      Barcode : String;
   END_VAR
   VAR_OUTPUT
      Ready : Bool;
      Running : Bool;
      Done : Bool;
      Valid : Bool;
      Barcode_Out : String;
      "Counter" : UInt;
   END_VAR
   VAR
      State : UInt;
      R_TRIG_Instance { S7_SetPoint := 'True'} : R_TRIG;
      IEC_Timer_0_Instance { S7_SetPoint := 'True'} : TON_TIME;
      IEC_Timer_0_Instance_1 { S7_SetPoint := 'True'} : TP_TIME;
   END_VAR
BEGIN
   #R_TRIG_Instance(CLK:=#Start);

   IF #R_TRIG_Instance.Q THEN
       IF #State = 0 THEN
           #State := 10;
       END_IF;
   END_IF;

   CASE #State OF

       0: // IDLE
           #Running := FALSE;
           #Ready := TRUE;
           #IEC_Timer_0_Instance(IN := FALSE,
                                 PT := T#0S);
           "IEC_Timer_0_DB_19".TP(IN := FALSE,
                                  PT := T#0S);

       10: // Start
           #Barcode_Out := '';
           #Done := FALSE;
           #Valid := FALSE;
           #Ready := FALSE;
           #Running := TRUE;
           #State := 20;

       20: // Reading code
           "Control_DB".InBarcode_Station.Start := FALSE;
           "Control_DB".InBarcode_Station."Reading Gate number" := "FindStringField"(FieldName := 'Number', JsonStr := "SICK_Barcode_DB".Result);
           "Control_DB".Inbound_Cnv.Inputs.Barcode := "FindStringField"(FieldName := 'Code', JsonStr := "SICK_Barcode_DB".Result);
           "Control_DB".InBarcode_Station."Number of Reading Gates" := "FindStringField"(FieldName := 'NRG', JsonStr := "SICK_Barcode_DB".Result);
           "Auto_Start_Barcode" := TRUE;

           //Check if the gate is open
               IF "Control_DB".InBarcode_Station."Number of Reading Gates" <> "Control_DB".InBarcode_Station."Number of Reading Gates OLD" THEN
                   "Control_DB".InBarcode_Station."Number of Reading Gates OLD" := "Control_DB".InBarcode_Station."Number of Reading Gates";
               END_IF;

               //Timer to read the barcode
               #IEC_Timer_0_Instance(IN := TRUE,
                                     PT := T#7S);

               //If a new code was read or the time finished
               IF "Control_DB".InBarcode_Station."Reading Gate number" <> "Control_DB".InBarcode_Station."Reading Gate number OLD" OR #IEC_Timer_0_Instance.Q THEN
                   "Auto_Start_Barcode" := FALSE; //Close the gate
                   //New code
                   IF "Control_DB".InBarcode_Station."Reading Gate number" <> "Control_DB".InBarcode_Station."Reading Gate number OLD" THEN
                       //Check if the string is not empty
                       IF LEN(IN := "SICK_Barcode_DB".Result) > 1 AND "Control_DB".InBarcode_Station."Reading Gate number" <> '' THEN
                           #Valid := TRUE;
                           #Barcode_Out := "Control_DB".Inbound_Cnv.Inputs.Barcode;
                       ELSE //Empty
                           #Valid := FALSE;
                           #Barcode_Out := '';
                       END_IF;
                       //Save OLD
                       "Control_DB".InBarcode_Station."Reading Gate number OLD" := "Control_DB".InBarcode_Station."Reading Gate number";
                       #IEC_Timer_0_Instance(IN := FALSE,
                                             PT := T#0S);
                           #State := 30;
                       ELSE // No code
                       #Valid := FALSE;
                       #Barcode_Out := '';
                       #IEC_Timer_0_Instance(IN := FALSE,
                                             PT := T#0S);
                       #State := 30;
                   END_IF;
               END_IF;

           30: // Finally
               "IEC_Timer_0_DB_19".TP(IN := FALSE,
                                      PT := T#0S);
               "Auto_Stop_Barcode" := TRUE; //Close gate
               //Make sure the command was sent
               IF "Auto_Stop_Barcode" THEN
                   #Counter := #Counter + 1;
                   #Running := FALSE;
                   #Done := TRUE;
                   #State := 0;
               END_IF;
   END_CASE;
END_FUNCTION_BLOCK

FUNCTION_BLOCK "Stack_Lights"   // FB21, SCL
{ S7_Optimized_Access := 'TRUE' }
VERSION : 0.1
// stored: AutoNumber true, IsIECCheckEnabled false, IsRetainMemResEnabled false, MemoryReserve 100, SetENOAutomatically false, UDAEnableTagReadback false
   VAR_INPUT
      VTD_Mode : UInt;
      Fault : Bool;
   END_VAR
   VAR_OUTPUT
      Red : Bool;
      Green : Bool;
      Blue : Bool;
      Buzzer : Bool;
   END_VAR
BEGIN
   //Commands for Stack Light

   IF #VTD_Mode = 1 THEN  // (1)Manual = Yellow
       #Blue := TRUE;
       #Red := TRUE;
       #Green := FALSE;
   ELSIF #VTD_Mode = 2 THEN  // (2)Semi-Auto = Blue
       #Green := FALSE;
       #Blue := TRUE;
       #Red := FALSE;
   ELSIF #VTD_Mode = 3 THEN  // (3)Auto = Green
       #Green := TRUE;
       #Red := FALSE;
       #Blue := FALSE;
   ELSIF #Fault THEN  // Fault = Red
       #Red := TRUE;
       #Green := FALSE;
       #Blue := FALSE;
   ELSE
       #Green := FALSE;
       #Red := FALSE;
       #Blue := FALSE;
   END_IF;
END_FUNCTION_BLOCK

